                       80: //Check which conveyor
                           //Popup 2 conveyor to popup conveyor 3
                           IF #Source_Location_Carousel.Device_Type = 16 AND #Destination_Location_Carousel.Device_Type = 17 AND "Control_DB".PopUp_Cnv[2].Cnv_Occupied AND
                               NOT "Control_DB".PopUp_Cnv[3].Cnv_Occupied AND "Control_DB".PopUp_Cnv[2].Inputs."Lift Down" AND "Control_DB".PopUp_Cnv[3].Inputs."Lift Down"
                           THEN //All good
                               "Control_DB"."Carrousel_Order Table".SM_State := "Control_DB".PopUp_Cnv[3].SM_State;
                               #State_Carrousel := 100;// Chain Transfer
                           ELSIF #Source_Location_Carousel.Device_Type = 16 AND #Destination_Location_Carousel.Device_Type = 17 AND "Control_DB".PopUp_Cnv[2].Cnv_Occupied AND
                               NOT "Control_DB".PopUp_Cnv[3].Cnv_Occupied AND (NOT "Control_DB".PopUp_Cnv[2].Inputs."Lift Down" OR NOT "Control_DB".PopUp_Cnv[3].Inputs."Lift Down")
                           THEN //Lift
                               "Control_DB"."Carrousel_Order Table".SM_State := "Control_DB".PopUp_Cnv[3].SM_State;
                               #State_Carrousel := 90;// Lift pop up 2 OR 3 
                           END_IF;

                       90:  //Lift PopUps
                               "Control_DB"."Carrousel_Order Table".SM_State := "Control_DB".PopUp_Cnv[3].SM_State;
                               "Control_DB".PopUp_Cnv[2].Instruction.Lift_Down := NOT "Control_DB".PopUp_Cnv[2].Running AND NOT "Control_DB".PopUp_Cnv[2].Inputs."Lift Down";
                               "Control_DB".PopUp_Cnv[3].Instruction.Lift_Down := NOT "Control_DB".PopUp_Cnv[3].Running AND NOT "Control_DB".PopUp_Cnv[3].Inputs."Lift Down";
                               IF "Control_DB".PopUp_Cnv[2].Inputs."Lift Down" AND "Control_DB".PopUp_Cnv[3].Inputs."Lift Down" THEN
                                   #State_Carrousel := 100;
                               END_IF;

                           100: //Start the transfer
                           //Popup 2 to popup 3 conveyors
                                   "Control_DB".PopUp_Cnv[2].Instruction.Transfer_To_ID := "Settings_DB".PopUp_Cnv_Settings[3].ID;
                               "Control_DB"."Carrousel_Order Table".SM_State := "Control_DB".PopUp_Cnv[3].SM_State;//Current machine state
                               "Control_DB".PopUp_Cnv[3].Instruction.Start_Transfer := NOT "Control_DB".PopUp_Cnv[3].Running;
                               "Control_DB".PopUp_Cnv[2].Instruction.Start_Transfer := NOT "Control_DB".PopUp_Cnv[2].Running;
                               IF "Control_DB".PopUp_Cnv[3].Running AND "Control_DB".PopUp_Cnv[2].Running THEN
                                   "Control_DB"."Carrousel_Order Table".Movement_Ready := TRUE;
                                   //"Control_DB"."Carrousel_Order Table".Task_Data_Available := FALSE;
                                   #State_Carrousel := 110;
                               END_IF;

                       110: //Wait for the transfer to complete
                           //Popup 2 to popup 3 conveyors
                           "Control_DB"."Carrousel_Order Table".SM_State := "Control_DB".PopUp_Cnv[3].SM_State;
                           IF "Control_DB".PopUp_Cnv[3].Done AND "Control_DB".PopUp_Cnv[2].Done
                           THEN
                               "Control_DB"."Carrousel_Order Table".Movement_Request_Complete := TRUE;
                               #State_Carrousel := 120;
                           END_IF;

                       120: //Wait for the ACK before we go back to Idle
                           "Control_DB"."Carrousel_Order Table".SM_State := "Control_DB".PopUp_Cnv[3].SM_State;
                           IF "Control_DB"."Carrousel_Order Table".Movement_Request_Complete_Ack THEN
                               #State_Carrousel := 250;
                           END_IF;

                           //=========================== Transfer to pick station (From Pop Conveyor 4)  ===========================

                       130: //Check which conveyor
                               //Pop conveyor 4 to popup conveyor 1 (Pick Station)    
                           IF #Source_Location_Carousel.Device_Type = 18 AND #Destination_Location_Carousel.Device_Type = 41 AND "Control_DB".PopUp_Cnv[4].Cnv_Occupied AND
                               "Pick Station" AND "Control_DB".PopUp_Cnv[4].Inputs."Lift Down" AND "Control_DB".PopUp_Cnv[1].Inputs."Lift Down"
                           THEN //All good
                               "Control_DB"."Carrousel_Order Table".SM_State := "Control_DB".PopUp_Cnv[1].SM_State;
                               #State_Carrousel := 150;// Chain Transfer
                           ELSIF #Source_Location_Carousel.Device_Type = 18 AND #Destination_Location_Carousel.Device_Type = 41 AND "Control_DB".PopUp_Cnv[4].Cnv_Occupied AND
                               "Pick Station" AND (NOT "Control_DB".PopUp_Cnv[4].Inputs."Lift Down" OR NOT "Control_DB".PopUp_Cnv[1].Inputs."Lift Down")
                           THEN //Lift
                               "Control_DB"."Carrousel_Order Table".SM_State := "Control_DB".PopUp_Cnv[1].SM_State;
                               #State_Carrousel := 140;// Lift pop up 1
                           END_IF;

                       140:  //Lift PopUp
                           "Control_DB"."Carrousel_Order Table".SM_State := "Control_DB".PopUp_Cnv[1].SM_State;
                            // "Control_DB".PopUp_Cnv[1].Instruction.Lift_Down := NOT "Control_DB".PopUp_Cnv[1].Running AND NOT "Control_DB".PopUp_Cnv[1].Inputs."Lift Down";
                            "Control_DB".PopUp_Cnv[4].Instruction.Lift_Down := NOT "Control_DB".PopUp_Cnv[4].Running AND NOT "Control_DB".PopUp_Cnv[4].Inputs."Lift Down" ;
                            IF (*"Control_DB".PopUp_Cnv[1].Inputs."Lift Down" AND*) "Control_DB".PopUp_Cnv[4].Inputs."Lift Down" THEN
                                   #State_Carrousel := 150;
                               END_IF;

                       150: //Start the transfer
                           //Popup 4 TO Pick station conveyors
                               "Control_DB"."Carrousel_Order Table".SM_State := "Control_DB".PopUp_Cnv[1].SM_State;//Current machine state
                               "Control_DB".PopUp_Cnv[1].Instruction.Start_Transfer := NOT "Control_DB".PopUp_Cnv[1].Running;
                               IF "Control_DB".PopUp_Cnv[1].Running THEN
                                   "Control_DB"."Carrousel_Order Table".Movement_Ready := TRUE;
                                  // "Control_DB"."Carrousel_Order Table".Task_Data_Available := FALSE;
                                   #State_Carrousel := 160;
                               END_IF;

                       160: //Wait for the transfer to complete
                           //Popup 4 TO Pick station conveyors
                           "Control_DB"."Carrousel_Order Table".SM_State := "Control_DB".PopUp_Cnv[1].SM_State;
                           IF #Source_Location_Carousel.Device_Type = 18 AND #Destination_Location_Carousel.Device_Type = 41 AND
                               "Control_DB".PopUp_Cnv[1].Done
                           THEN
                               "Control_DB"."Carrousel_Order Table".Movement_Request_Complete := TRUE;
                               #State_Carrousel := 170;
                           END_IF;

                       170: //Wait for the ACK before we go back to Idle
                           "Control_DB"."Carrousel_Order Table".SM_State := "Control_DB".PopUp_Cnv[1].SM_State;
                           IF "Control_DB"."Carrousel_Order Table".Movement_Request_Complete_Ack THEN
                               #State_Carrousel := 250;
                           END_IF;

                           //=========================== Transfer from Pick station (To Pop Conveyor 1)  ===========================

                       180: //Check which conveyor
                               //Pick to popup conveyor 1   
                           IF #Source_Location_Carousel.Device_Type = 41 AND #Destination_Location_Carousel.Device_Type = 15 AND NOT "Pick Station" AND
                               NOT "Control_DB".PopUp_Cnv[1].Cnv_Occupied AND "Control_DB".PopUp_Cnv[1].Inputs."Lift Down"
                           THEN //All good
                               "Control_DB"."Carrousel_Order Table".SM_State := "Control_DB".PopUp_Cnv[1].SM_State;
                               #State_Carrousel := 200;// Chain Transfer
                           ELSIF #Source_Location_Carousel.Device_Type = 41 AND #Destination_Location_Carousel.Device_Type = 15 AND NOT "Pick Station" AND
                               NOT "Control_DB".PopUp_Cnv[1].Cnv_Occupied AND NOT "Control_DB".PopUp_Cnv[1].Inputs."Lift Down"
                           THEN //Lift
                               "Control_DB"."Carrousel_Order Table".SM_State := "Control_DB".PopUp_Cnv[1].SM_State;
                               #State_Carrousel := 190;// Lift pop up 1
                           END_IF;

                       190:  //Lift PopUps
                           "Control_DB"."Carrousel_Order Table".SM_State := "Control_DB".PopUp_Cnv[1].SM_State;
                           "Control_DB".PopUp_Cnv[1].Instruction.Lift_Down := NOT "Control_DB".PopUp_Cnv[1].Running AND NOT "Control_DB".PopUp_Cnv[1].Inputs."Lift Down";
                           IF "Control_DB".PopUp_Cnv[1].Inputs."Lift Down" THEN
                               #State_Carrousel := 200;
                           END_IF;

                       200: //Start the transfer
                           //Pick station TO Popup 1 conveyors
                               "Control_DB"."Carrousel_Order Table".SM_State := "Control_DB".PopUp_Cnv[1].SM_State;//Current machine state
                               "Control_DB".PopUp_Cnv[1].Instruction.Start_Transfer := NOT "Control_DB".PopUp_Cnv[1].Running;
                               IF "Control_DB".PopUp_Cnv[1].Running AND NOT "Control_DB".PopUp_Cnv[1].Done THEN
                                   "Control_DB"."Carrousel_Order Table".Movement_Ready := TRUE;
                                   //"Control_DB"."Carrousel_Order Table".Task_Data_Available := FALSE;
                                   #State_Carrousel := 210;
                               END_IF;

                       210: //Wait for the transfer to complete
                           //Pick station TO PopUp 1 conveyors
                           "Control_DB"."Carrousel_Order Table".SM_State := "Control_DB".PopUp_Cnv[1].SM_State;
                           IF "Control_DB".PopUp_Cnv[1].Done THEN
                               "Control_DB"."Carrousel_Order Table".Movement_Request_Complete := TRUE;
                               #State_Carrousel := 220;
                           END_IF;

                       220: //Wait for the ACK before we go back to Idle
                           "Control_DB"."Carrousel_Order Table".SM_State := "Control_DB".PopUp_Cnv[1].SM_State;
                           IF "Control_DB"."Carrousel_Order Table".Movement_Request_Complete_Ack THEN
                               #State_Carrousel := 250;
                           END_IF;

                           //=========================== Weigh Pallet  ===========================
                       230:
                          // "Control_DB"."Carrousel_Order Table".Task_Data_Available := FALSE;
                           "Control_DB"."Weighing Station".Start := TRUE;
                           "Control_DB"."Carrousel_Order Table".Movement_Ready := TRUE;
                           "Control_DB"."Carrousel_Order Table".SM_State := INT_TO_UINT("State_WS");
                           //Lift PopUp 1
                           "Control_DB".PopUp_Cnv[1].Instruction.Lift_Up := NOT "Control_DB".PopUp_Cnv[1].Running AND NOT "Control_DB".PopUp_Cnv[1].Inputs."Lift Up";

                           "IEC_Timer_0_DB_9".TON(IN:="Control_DB".PopUp_Cnv[1].Inputs."Lift Up",
                                                  PT:=T#500MS);
                           IF "IEC_Timer_0_DB_9".Q THEN
                               "Control_DB"."Weighing Station".Start := fALSE;
                               "IEC_Timer_0_DB_9".TON(IN := fALSE,
                                                      PT := T#0MS);
                               #State_Carrousel := 232;
                           END_IF;

                       232:
                           "Control_DB"."Carrousel_Order Table".SM_State := INT_TO_UINT("State_WS");
                           IF "Control_DB"."Weighing Station".Done THEN
                               "Control_DB"."Carrousel_Order Table".Movement_Request_Complete := TRUE;
                               IF "Control_DB"."Carrousel_Order Table".Movement_Request_Complete_Ack THEN
                                   #State_Carrousel := 250;
                               END_IF;
                           ELSE
                               #State_Carrousel := 250;
                           END_IF;

                           //=========================== Reset and Error States ===========================
                           250: //Reset all variable and return to idle

                           //Reset the OPC control variables
                               "Control_DB"."Carrousel_Order Table".SM_State := 0;
                               "Control_DB"."Carrousel_Order Table".Movement_Ready := FALSE;
                               "Control_DB"."Carrousel_Order Table".Movement_Request_Complete := FALSE;
                               "Control_DB"."Carrousel_Order Table".Movement_Request_Complete_Ack := FALSE;
                               "Control_DB"."Carrousel_Order Table".Task_Metadata := '';

                               "Control_DB"."Carrousel_Order Table".Task_Data_Available := FALSE; // Send the Task Data Available from WCS 
                               "Control_DB"."Carrousel_Order Table".Task_Type := 0; //  Send the Task Type - Roller to Roller Conveyor = Task Type = 6
                               "Control_DB"."Carrousel_Order Table".Task_ID := 0; // Send the Task ID number;
                               "Control_DB"."Carrousel_Order Table".Source_Location := 0; // Send the Source Location from the Conveyor
                               "Control_DB"."Carrousel_Order Table".Destination_Location := 0; // Send the Destination Location 
                               #Destination_Location_Carousel.Device_Type:=0;
                               #Source_Location_Carousel.Device_Type := 0;

                           //Reset conveyor variables
                           "Control_DB".Inbound_Cnv.Instruction.Start_Transfer := FALSE;
                           "Control_DB".Inbound_Cnv.Instruction.Task_ID := 0;
                           "Control_DB".Inbound_Cnv.Instruction.Task_Metadata := '';
                           "Control_DB".Inbound_Cnv.Current_Task_Type := 0;
                           "Control_DB".Inbound_Cnv.Instruction.Transfer_From_ID := 0;
                           "Control_DB".Inbound_Cnv.Instruction.Transfer_To_ID := 0;

                           "Control_DB".Outbound_Cnv.Instruction.Start_Transfer := FALSE;
                           "Control_DB".Outbound_Cnv.Instruction.Task_ID := 0;
                           "Control_DB".Outbound_Cnv.Instruction.Task_Metadata := '';
                           "Control_DB".Outbound_Cnv.Current_Task_Type := 0;
                           "Control_DB".Outbound_Cnv.Instruction.Transfer_From_ID := 0;
                           "Control_DB".Outbound_Cnv.Instruction.Transfer_To_ID := 0;

                           FOR #i := 1 TO 4 DO
                               "Control_DB".PopUp_Cnv[#i].Instruction.Start_Transfer := FALSE;
                               "Control_DB".PopUp_Cnv[#i].Instruction.Task_ID := 0;
                               "Control_DB".PopUp_Cnv[#i].Instruction.Task_Metadata := '';
                               "Control_DB".PopUp_Cnv[#i].Current_Task_Type := 0;
                               "Control_DB".PopUp_Cnv[#i].Instruction.Transfer_From_ID := 0;
                               "Control_DB".PopUp_Cnv[#i].Instruction.Transfer_To_ID := 0;
                           END_FOR;

                           "Error_Word_1".%X1 := FALSE;

                           #State_Carrousel := 0;

                           400:// Error state
                               "Control_DB"."Carrousel_Order Table".Task_Metadata := '';
                               "Control_DB"."Carrousel_Order Table".Task_Data_Available := FALSE; // Send the Task Data Available from WCS 
                               "Control_DB"."Carrousel_Order Table".Task_Type := 0; //  Send the Task Type - Roller to Roller Conveyor = Task Type = 6
                               "Control_DB"."Carrousel_Order Table".Task_ID := 0; // Send the Task ID number;
                               "Control_DB"."Carrousel_Order Table".Source_Location := 0; // Send the Source Location from the Conveyor
                               "Control_DB"."Carrousel_Order Table".Destination_Location := 0; // Send the Destination Location

                               #Destination_Location_Carousel.Device_Type := 0;
                               #Source_Location_Carousel.Device_Type := 0;


                           IF "Control_DB".VTD_Control.Instruction.Reset
                           THEN
                               #State_Carrousel := 250;
                           END_IF;

                       ELSE
                           ;
                   END_CASE;
                   ELSIF "Carrousel_In_Automatic" AND NOT #OPC_Enable THEN
                       "Control_DB"."Carrousel_Order Table".Task_Metadata := '';
                       //Reset all variable and return to idle

                       //Reset the OPC control variables
                       "Control_DB"."Carrousel_Order Table".SM_State := 0;
                       "Control_DB"."Carrousel_Order Table".Movement_Ready := FALSE;
                       "Control_DB"."Carrousel_Order Table".Movement_Request_Complete := FALSE;

                       "Control_DB"."Carrousel_Order Table".Task_Data_Available := FALSE; // Send the Task Data Available from WCS 
                       "Control_DB"."Carrousel_Order Table".Task_Type := 0; //  Send the Task Type - Roller to Roller Conveyor = Task Type = 6
                       "Control_DB"."Carrousel_Order Table".Task_ID := 0; // Send the Task ID number;
                       "Control_DB"."Carrousel_Order Table".Source_Location := 0; // Send the Source Location from the Conveyor
                       "Control_DB"."Carrousel_Order Table".Destination_Location := 0; // Send the Destination Location

                       #Destination_Location_Carousel.Device_Type := 0;
                       #Source_Location_Carousel.Device_Type := 0;

                       //Reset conveyor variables
                       "Control_DB".Inbound_Cnv.Instruction.Start_Transfer := FALSE;
                       "Control_DB".Inbound_Cnv.Instruction.Task_ID := 0;
                       "Control_DB".Inbound_Cnv.Instruction.Task_Metadata := '';//
                       "Control_DB".Inbound_Cnv.Instruction.Transfer_From_ID := 0;
                       "Control_DB".Inbound_Cnv.Instruction.Transfer_To_ID := 0;

                       "Control_DB".Outbound_Cnv.Instruction.Start_Transfer := FALSE;
                       "Control_DB".Outbound_Cnv.Instruction.Task_ID := 0;
                       "Control_DB".Outbound_Cnv.Instruction.Task_Metadata := '';//
                       "Control_DB".Outbound_Cnv.Instruction.Transfer_From_ID := 0;
                       "Control_DB".Outbound_Cnv.Instruction.Transfer_To_ID := 0;

                       FOR #i := 1 TO 4 DO
                           "Control_DB".PopUp_Cnv[#i].Instruction.Start_Transfer := FALSE;
                           "Control_DB".PopUp_Cnv[#i].Instruction.Task_ID := 0;
                           "Control_DB".PopUp_Cnv[#i].Instruction.Task_Metadata := '';
                           "Control_DB".PopUp_Cnv[#i].Current_Task_Type := 0;
                           "Control_DB".PopUp_Cnv[#i].Instruction.Transfer_From_ID := 0;
                           "Control_DB".PopUp_Cnv[#i].Instruction.Transfer_To_ID := 0;
                       END_FOR;
                   END_IF;
       END_REGION
   END_REGION

   REGION SHUTTLES POSITION
       FOR #f := 1 TO "Settings_DB".System_Settings.Shuttle_Count DO
           "Control_DB".Shuttles_Position[#f].x := "Shuttle_MQTT_DB".Shuttle_MQTT[#f].Message.Shuttle_Status.Position_X;
           "Control_DB".Shuttles_Position[#f].y := "Shuttle_MQTT_DB".Shuttle_MQTT[#f].Message.Shuttle_Status.Position_Y;
       END_FOR;
   END_REGION

   REGION SM STATE MAESTRO
       // Statement section - Send the State machine to Maestro "Emulating" openTCS states
       // 
      // // "Control_DB".WMS_OPC_UA.SM_State_Maestro; // State to send Devices to Maestro
      //  IF #State_VTD = 0 THEN

      //      "Control_DB"."VTD_Order Table".SM_State_Maestro := 0;//"LIMBO" condition 

      //  ELSIF "Control_DB"."VTD_Order Table".SM_State = 10 THEN
      //      ;
      //      // "Control_DB".WMS_OPC_UA.SM_State_Maestro := 1;//RAW conidtion => Maestro will write this condition

      //      //////////////////////////////////////////////////////////////////////////////////////////////////////////////////////      
      //      // QUEUED ANY DEVICE    
      //  // ELSIF "Control_DB".WMS_OPC_UA.Task_Data_Available AND #State >= 10 AND #State <= 20 THEN
      //  ELSIF "Control_DB"."VTD_Order Table".Task_Data_Available AND NOT "Control_DB"."VTD_Order Table".Movement_Ready AND "Control_DB"."VTD_Order Table".SM_State_Maestro = 1 THEN
      //      "Control_DB"."VTD_Order Table".SM_State_Maestro := 2;//QUEUED condition =>ANY device (Conveyor, VTD OR Shuttle)  

      //      //////////////////////////////////////////////////////////////////////////////////////////////////////////////////////       
      //      // Any Device RUNNING on the system (VTD - Conveyor Transfer - Shuttle Transfer) 
      //  ELSIF ("Control_DB"."VTD_Order Table".Task_Type = 4 OR "Control_DB"."VTD_Order Table".Task_Type = 5
      //      OR "Control_DB"."VTD_Order Table".Task_Type = 1 OR "Control_DB"."VTD_Order Table".Task_Type = 2 OR "Control_DB"."VTD_Order Table".Task_Type = 3)
      //      AND "Control_DB"."VTD_Order Table".Movement_Ready AND NOT "Control_DB"."VTD_Order Table".Movement_Request_Complete THEN

      //      "Control_DB"."VTD_Order Table".SM_State_Maestro := 3;//RUNNING condition

      //      // Any Device DONE on the system (VTD - Coneveyor Transfer - Shuttle Transfer) 
      //  ELSIF ("Control_DB"."VTD_Order Table".Task_Type = 4 OR "Control_DB"."VTD_Order Table".Task_Type = 5
      //      OR "Control_DB"."VTD_Order Table".Task_Type = 1 OR "Control_DB"."VTD_Order Table".Task_Type = 2 OR "Control_DB"."VTD_Order Table".Task_Type = 3)
      //      AND (*"Control_DB".WMS_OPC_UA.Movement_Request_Complete AND "Control_DB".WMS_OPC_UA.Movement_Ready*)#State_VTD = 120 OR #State_VTD = 45 OR #State_VTD = 90 THEN

      //      "Control_DB"."VTD_Order Table".SM_State_Maestro := 4;//DONE condition

      //      // Any Device ERRORS on the system (VTD - Coneveyor Transfer - Shuttle Transfer)  
      //  ELSIF ("Control_DB"."VTD_Order Table".Task_Type = 4 OR "Control_DB"."VTD_Order Table".Task_Type = 5
      //      OR "Control_DB"."VTD_Order Table".Task_Type = 1 OR "Control_DB"."VTD_Order Table".Task_Type = 2 OR "Control_DB"."VTD_Order Table".Task_Type = 3)
      //      AND "Control_DB"."VTD_Order Table".SM_State = 400 THEN

      //      "Control_DB"."VTD_Order Table".SM_State_Maestro := 5;//ERROR condition => Conveyors   
      //  END_IF;
      //      /////////////////////////////////////////////////////////////////////////////////////////////        



       // "Control_DB".WMS_OPC_UA.SM_State_Maestro; // State to send Devices to Maestro
        IF #State_VTD = 0 THEN
            ;
            //"System_DB_VTD".OrderTable[1].OPC_Control.SM_State_Maestro := 0;//"LIMBO" condition 

        ELSIF "Control_DB"."VTD_Order Table".SM_State = 10 THEN
            ;
            // "Control_DB".WMS_OPC_UA.SM_State_Maestro := 1;//RAW conidtion => Maestro will write this condition

            //////////////////////////////////////////////////////////////////////////////////////////////////////////////////////      
            // QUEUED ANY DEVICE    
        // ELSIF "Control_DB".WMS_OPC_UA.Task_Data_Available AND #State >= 10 AND #State <= 20 THEN
        ELSIF "Control_DB"."VTD_Order Table".Task_Data_Available AND NOT "Control_DB"."VTD_Order Table".Movement_Ready AND "System_DB_VTD".OrderTable[1].OPC_Control.SM_State_Maestro = 1 THEN
            "System_DB_VTD".OrderTable[1].OPC_Control.SM_State_Maestro := 2;//QUEUED condition =>ANY device (Conveyor, VTD OR Shuttle)  

            //////////////////////////////////////////////////////////////////////////////////////////////////////////////////////       
            // Any Device RUNNING on the system (VTD - Conveyor Transfer - Shuttle Transfer) 
        ELSIF ("Control_DB"."VTD_Order Table".Task_Type = 4 OR "Control_DB"."VTD_Order Table".Task_Type = 5
            OR "Control_DB"."VTD_Order Table".Task_Type = 1 OR "Control_DB"."VTD_Order Table".Task_Type = 2 OR "Control_DB"."VTD_Order Table".Task_Type = 3)
            AND "Control_DB"."VTD_Order Table".Movement_Ready AND NOT "Control_DB"."VTD_Order Table".Movement_Request_Complete THEN

            "System_DB_VTD".OrderTable[1].OPC_Control.SM_State_Maestro  := 3;//RUNNING condition

            // Any Device DONE on the system (VTD - Coneveyor Transfer - Shuttle Transfer) 
        ELSIF ("Control_DB"."VTD_Order Table".Task_Type = 4 OR "Control_DB"."VTD_Order Table".Task_Type = 5
            OR "Control_DB"."VTD_Order Table".Task_Type = 1 OR "Control_DB"."VTD_Order Table".Task_Type = 2 OR "Control_DB"."VTD_Order Table".Task_Type = 3)
            AND (*"Control_DB".WMS_OPC_UA.Movement_Request_Complete AND "Control_DB".WMS_OPC_UA.Movement_Ready*)#State_VTD = 120 OR #State_VTD = 45 OR #State_VTD = 90 THEN

            "System_DB_VTD".OrderTable[1].OPC_Control.SM_State_Maestro := 4;//DONE condition

            // Any Device ERRORS on the system (VTD - Coneveyor Transfer - Shuttle Transfer)  
        ELSIF ("Control_DB"."VTD_Order Table".Task_Type = 4 OR "Control_DB"."VTD_Order Table".Task_Type = 5
            OR "Control_DB"."VTD_Order Table".Task_Type = 1 OR "Control_DB"."VTD_Order Table".Task_Type = 2 OR "Control_DB"."VTD_Order Table".Task_Type = 3)
            AND "Control_DB"."VTD_Order Table".SM_State = 400 THEN

            "System_DB_VTD".OrderTable[1].OPC_Control.SM_State_Maestro := 5;//ERROR condition => Conveyors   
        END_IF;
            /////////////////////////////////////////////////////////////////////////////////////////////        


      //  //     //////////////////////////////////////////////////////////////////////////////////////////////////////////////////////       
      //  //     // Any VTD RUNNING on the system (VTD) 
      //  // ELSIF "Control_DB".WMS_OPC_UA.Task_Type = 1
      //  //     AND "Control_DB".WMS_OPC_UA.SM_State >= 35 AND "Control_DB".WMS_OPC_UA.SM_State < 100 AND #State > 20 THEN

      //  //     "Control_DB".WMS_OPC_UA.SM_State_Maestro := 3;//RUNNING condition => VTD

      //  //     // Any VTD DONE on the system (VTD) 
      //  // ELSIF "Control_DB".WMS_OPC_UA.Task_Type = 1
      //  //     AND "Control_DB".WMS_OPC_UA.SM_State = 100 AND #State > 20 THEN

      //  //     "Control_DB".WMS_OPC_UA.SM_State_Maestro := 4;//DONE condition => VTD

      //  //     // Any VTD ERRORS on the system (VTD) 
      //  // ELSIF "Control_DB".WMS_OPC_UA.Task_Type = 1
      //  //     AND "Control_DB".WMS_OPC_UA.SM_State = 400 THEN

      //  //     "Control_DB".WMS_OPC_UA.SM_State_Maestro := 5;//ERROR condition => VTD   



      //  //     //////////////////////////////////////////////////////////////////////////////////////////////////////////////////////       
      //  //     // Any Shuttle Interlock RUNNING on the system (Shuttle) 
      //  // ELSIF "Control_DB".WMS_OPC_UA.Task_Type = 2 OR "Control_DB".WMS_OPC_UA.Task_Type = 3
      //  //     AND "Control_DB".WMS_OPC_UA.SM_State >= 35 AND "Control_DB".WMS_OPC_UA.SM_State < 100 AND #State > 20 THEN

      //  //     "Control_DB".WMS_OPC_UA.SM_State_Maestro := 3;//RUNNING condition => Shuttle

      //  //     // Any Shuttle Interlock  DONE on the system (Shuttle) 
      //  // ELSIF "Control_DB".WMS_OPC_UA.Task_Type = 2 OR "Control_DB".WMS_OPC_UA.Task_Type = 3
      //  //     AND "Control_DB".WMS_OPC_UA.SM_State = 100 AND #State > 20 THEN

      //  //     "Control_DB".WMS_OPC_UA.SM_State_Maestro := 4;//DONE condition => Shuttle

      //  //     // Any Shuttle Interlock ERRORS on the system (Shuttle) 
      //  // ELSIF "Control_DB".WMS_OPC_UA.Task_Type = 2 OR "Control_DB".WMS_OPC_UA.Task_Type = 3
      //  //     AND "Control_DB".WMS_OPC_UA.SM_State = 400 THEN

      //  //     "Control_DB".WMS_OPC_UA.SM_State_Maestro := 5;//ERROR condition => Shuttle          

      //  // END_IF;


       // // "Control_DB".WMS_OPC_UA.SM_State_Maestro; // State to send Devices to Maestro
       //  IF #State_VTD = 0 THEN

       //      "Control_DB"."VTD_Order Table".SM_State_Maestro := 0;//"LIMBO" condition 

       //  ELSIF "Control_DB"."VTD_Order Table".SM_State = 10 THEN
       //      ;
       //      // "Control_DB".WMS_OPC_UA.SM_State_Maestro := 1;//RAW conidtion => Maestro will write this condition

       //      //////////////////////////////////////////////////////////////////////////////////////////////////////////////////////      
       //      // QUEUED ANY DEVICE    
       //  // ELSIF "Control_DB".WMS_OPC_UA.Task_Data_Available AND #State >= 10 AND #State <= 20 THEN
       //  ELSIF "Control_DB"."VTD_Order Table".Task_Data_Available AND NOT "Control_DB"."VTD_Order Table".Movement_Ready AND "Control_DB"."VTD_Order Table".SM_State_Maestro = 1 THEN
       //      "Control_DB"."VTD_Order Table".SM_State_Maestro := 2;//QUEUED condition =>ANY device (Conveyor, VTD OR Shuttle)  

       //      //////////////////////////////////////////////////////////////////////////////////////////////////////////////////////       
       //      // Any Device RUNNING on the system (VTD - Conveyor Transfer - Shuttle Transfer) 
       //  ELSIF ("Control_DB"."VTD_Order Table".Task_Type = 4 OR "Control_DB"."VTD_Order Table".Task_Type = 5
       //      OR "Control_DB"."VTD_Order Table".Task_Type = 1 OR "Control_DB"."VTD_Order Table".Task_Type = 2 OR "Control_DB"."VTD_Order Table".Task_Type = 3)
       //      AND "Control_DB"."VTD_Order Table".Movement_Ready AND NOT "Control_DB"."VTD_Order Table".Movement_Request_Complete THEN

       //      "Control_DB"."VTD_Order Table".SM_State_Maestro := 3;//RUNNING condition

       //      // Any Device DONE on the system (VTD - Coneveyor Transfer - Shuttle Transfer) 
       //  ELSIF ("Control_DB"."VTD_Order Table".Task_Type = 4 OR "Control_DB"."VTD_Order Table".Task_Type = 5
       //      OR "Control_DB"."VTD_Order Table".Task_Type = 1 OR "Control_DB"."VTD_Order Table".Task_Type = 2 OR "Control_DB"."VTD_Order Table".Task_Type = 3)
       //      AND (*"Control_DB".WMS_OPC_UA.Movement_Request_Complete AND "Control_DB".WMS_OPC_UA.Movement_Ready*)#State_VTD = 120 OR #State_VTD = 45 OR #State_VTD = 90 THEN

       //      "Control_DB"."VTD_Order Table".SM_State_Maestro := 4;//DONE condition

       //      // Any Device ERRORS on the system (VTD - Coneveyor Transfer - Shuttle Transfer)  
       //  ELSIF ("Control_DB"."VTD_Order Table".Task_Type = 4 OR "Control_DB"."VTD_Order Table".Task_Type = 5
       //      OR "Control_DB"."VTD_Order Table".Task_Type = 1 OR "Control_DB"."VTD_Order Table".Task_Type = 2 OR "Control_DB"."VTD_Order Table".Task_Type = 3)
       //      AND "Control_DB"."VTD_Order Table".SM_State = 400 THEN

       //      "Control_DB"."VTD_Order Table".SM_State_Maestro := 5;//ERROR condition => Conveyors   
       //  END_IF;
       //      /////////////////////////////////////////////////////////////////////////////////////////////        

       //  //     //////////////////////////////////////////////////////////////////////////////////////////////////////////////////////       
       //  //     // Any VTD RUNNING on the system (VTD) 
       //  // ELSIF "Control_DB".WMS_OPC_UA.Task_Type = 1
       //  //     AND "Control_DB".WMS_OPC_UA.SM_State >= 35 AND "Control_DB".WMS_OPC_UA.SM_State < 100 AND #State > 20 THEN

       //  //     "Control_DB".WMS_OPC_UA.SM_State_Maestro := 3;//RUNNING condition => VTD

       //  //     // Any VTD DONE on the system (VTD) 
       //  // ELSIF "Control_DB".WMS_OPC_UA.Task_Type = 1
       //  //     AND "Control_DB".WMS_OPC_UA.SM_State = 100 AND #State > 20 THEN

       //  //     "Control_DB".WMS_OPC_UA.SM_State_Maestro := 4;//DONE condition => VTD

       //  //     // Any VTD ERRORS on the system (VTD) 
       //  // ELSIF "Control_DB".WMS_OPC_UA.Task_Type = 1
       //  //     AND "Control_DB".WMS_OPC_UA.SM_State = 400 THEN

       //  //     "Control_DB".WMS_OPC_UA.SM_State_Maestro := 5;//ERROR condition => VTD   



       //  //     //////////////////////////////////////////////////////////////////////////////////////////////////////////////////////       
       //  //     // Any Shuttle Interlock RUNNING on the system (Shuttle) 
       //  // ELSIF "Control_DB".WMS_OPC_UA.Task_Type = 2 OR "Control_DB".WMS_OPC_UA.Task_Type = 3
       //  //     AND "Control_DB".WMS_OPC_UA.SM_State >= 35 AND "Control_DB".WMS_OPC_UA.SM_State < 100 AND #State > 20 THEN

       //  //     "Control_DB".WMS_OPC_UA.SM_State_Maestro := 3;//RUNNING condition => Shuttle

       //  //     // Any Shuttle Interlock  DONE on the system (Shuttle) 
       //  // ELSIF "Control_DB".WMS_OPC_UA.Task_Type = 2 OR "Control_DB".WMS_OPC_UA.Task_Type = 3
       //  //     AND "Control_DB".WMS_OPC_UA.SM_State = 100 AND #State > 20 THEN

       //  //     "Control_DB".WMS_OPC_UA.SM_State_Maestro := 4;//DONE condition => Shuttle

       //  //     // Any Shuttle Interlock ERRORS on the system (Shuttle) 
       //  // ELSIF "Control_DB".WMS_OPC_UA.Task_Type = 2 OR "Control_DB".WMS_OPC_UA.Task_Type = 3
       //  //     AND "Control_DB".WMS_OPC_UA.SM_State = 400 THEN

       //  //     "Control_DB".WMS_OPC_UA.SM_State_Maestro := 5;//ERROR condition => Shuttle          

       //  // END_IF;

   END_REGION


   REGION SM STATE MAESTRO - Carousel
       // Statement section - Send the State machine to Maestro "Emulating" openTCS states
       // 

       (*
       IF #State_Carrousel = 0 THEN

           "Control_DB"."Carrousel_Order Table".SM_State_Maestro := 0;//"LIMBO" condition 

       ELSIF "Control_DB"."Carrousel_Order Table".SM_State = 10 THEN
           ;
           // "Control_DB".WMS_OPC_UA.SM_State_Maestro := 1;//RAW conidtion => Maestro will write this condition

           //////////////////////////////////////////////////////////////////////////////////////////////////////////////////////      
           // QUEUED ANY DEVICE    
           // ELSIF "Control_DB".WMS_OPC_UA.Task_Data_Available AND #State >= 10 AND #State <= 20 THEN
       ELSIF "Control_DB"."Carrousel_Order Table".Task_Data_Available AND NOT "Control_DB"."Carrousel_Order Table".Movement_Ready AND "Control_DB"."Carrousel_Order Table".SM_State_Maestro = 1 THEN
           "Control_DB"."Carrousel_Order Table".SM_State_Maestro := 2;//QUEUED condition =>ANY device (Conveyor, VTD OR Shuttle)  

           //////////////////////////////////////////////////////////////////////////////////////////////////////////////////////       
           // Any Device RUNNING on the system (VTD - Conveyor Transfer - Shuttle Transfer) 
       ELSIF ("Control_DB"."Carrousel_Order Table".Task_Type = 6 OR "Control_DB"."Carrousel_Order Table".Task_Type = 7
           OR "Control_DB"."Carrousel_Order Table".Task_Type = 8 OR "Control_DB"."Carrousel_Order Table".Task_Type = 9
           OR "Control_DB"."Carrousel_Order Table".Task_Type = 10 OR "Control_DB"."Carrousel_Order Table".Task_Type = 14 OR "Control_DB"."Carrousel_Order Table".Task_Type = 16)
           AND "Control_DB"."Carrousel_Order Table".Movement_Ready AND NOT "Control_DB"."Carrousel_Order Table".Movement_Request_Complete THEN

           "Control_DB"."Carrousel_Order Table".SM_State_Maestro := 3;//RUNNING condition

           // Any Device DONE on the system (VTD - Coneveyor Transfer - Shuttle Transfer) 
       ELSIF ("Control_DB"."Carrousel_Order Table".Task_Type = 6 OR "Control_DB"."Carrousel_Order Table".Task_Type = 7
           OR "Control_DB"."Carrousel_Order Table".Task_Type = 8 OR "Control_DB"."Carrousel_Order Table".Task_Type = 9
           OR "Control_DB"."Carrousel_Order Table".Task_Type = 10 OR "Control_DB"."Carrousel_Order Table".Task_Type = 14 OR "Control_DB"."Carrousel_Order Table".Task_Type = 16)
           AND (*"Control_DB".WMS_OPC_UA.Movement_Request_Complete AND "Control_DB".WMS_OPC_UA.Movement_Ready*)#State_Carrousel = 70 OR #State_Carrousel = 120 OR #State_Carrousel = 170 OR #State_Carrousel = 220 OR #State_Carrousel = 232 THEN

           "Control_DB"."Carrousel_Order Table".SM_State_Maestro := 4;//DONE condition

           // Any Device ERRORS on the system (VTD - Coneveyor Transfer - Shuttle Transfer)  
       ELSIF ("Control_DB"."Carrousel_Order Table".Task_Type = 6 OR "Control_DB"."Carrousel_Order Table".Task_Type = 7
           OR "Control_DB"."Carrousel_Order Table".Task_Type = 8 OR "Control_DB"."Carrousel_Order Table".Task_Type = 9
           OR "Control_DB"."Carrousel_Order Table".Task_Type = 10 OR "Control_DB"."Carrousel_Order Table".Task_Type = 14 OR "Control_DB"."Carrousel_Order Table".Task_Type = 16)
           AND "Control_DB"."Carrousel_Order Table".SM_State = 400 THEN

           "Control_DB"."Carrousel_Order Table".SM_State_Maestro := 5;//ERROR condition => Conveyors   
       END_IF;
       /////////////////////////////////////////////////////////////////////////////////////////////        
       *)


       IF #State_Carrousel = 0 THEN
           ;
           //"Control_DB"."Carrousel_Order Table".SM_State_Maestro := 0;//"LIMBO" condition 
           //"System_DB_Carousel".OrderTable[1].OPC_Control.SM_State_Maestro := 0;

       ELSIF "Control_DB"."Carrousel_Order Table".SM_State = 10 THEN
           ;
           // "Control_DB".WMS_OPC_UA.SM_State_Maestro := 1;//RAW conidtion => Maestro will write this condition

           //////////////////////////////////////////////////////////////////////////////////////////////////////////////////////      
           // QUEUED ANY DEVICE    
           // ELSIF "Control_DB".WMS_OPC_UA.Task_Data_Available AND #State >= 10 AND #State <= 20 THEN
       ELSIF "Control_DB"."Carrousel_Order Table".Task_Data_Available AND NOT "Control_DB"."Carrousel_Order Table".Movement_Ready AND "System_DB_Carousel".OrderTable[1].OPC_Control.SM_State_Maestro = 1 THEN
           "System_DB_Carousel".OrderTable[1].OPC_Control.SM_State_Maestro := 2;//QUEUED condition =>ANY device (Conveyor, VTD OR Shuttle)  

           //////////////////////////////////////////////////////////////////////////////////////////////////////////////////////       
           // Any Device RUNNING on the system (VTD - Conveyor Transfer - Shuttle Transfer) 
       ELSIF ("Control_DB"."Carrousel_Order Table".Task_Type = 6 OR "Control_DB"."Carrousel_Order Table".Task_Type = 7
           OR "Control_DB"."Carrousel_Order Table".Task_Type = 8 OR "Control_DB"."Carrousel_Order Table".Task_Type = 9
           OR "Control_DB"."Carrousel_Order Table".Task_Type = 10 OR "Control_DB"."Carrousel_Order Table".Task_Type = 14 OR "Control_DB"."Carrousel_Order Table".Task_Type = 16)
           AND "Control_DB"."Carrousel_Order Table".Movement_Ready AND NOT "Control_DB"."Carrousel_Order Table".Movement_Request_Complete THEN

           "System_DB_Carousel".OrderTable[1].OPC_Control.SM_State_Maestro := 3;//RUNNING condition

           // Any Device DONE on the system (VTD - Coneveyor Transfer - Shuttle Transfer) 
       ELSIF ("Control_DB"."Carrousel_Order Table".Task_Type = 6 OR "Control_DB"."Carrousel_Order Table".Task_Type = 7
           OR "Control_DB"."Carrousel_Order Table".Task_Type = 8 OR "Control_DB"."Carrousel_Order Table".Task_Type = 9
           OR "Control_DB"."Carrousel_Order Table".Task_Type = 10 OR "Control_DB"."Carrousel_Order Table".Task_Type = 14 OR "Control_DB"."Carrousel_Order Table".Task_Type = 16)
           AND (*"Control_DB".WMS_OPC_UA.Movement_Request_Complete AND "Control_DB".WMS_OPC_UA.Movement_Ready*)#State_Carrousel = 70 OR #State_Carrousel = 120 OR #State_Carrousel = 170 OR #State_Carrousel = 220 OR #State_Carrousel = 232 THEN

           "System_DB_Carousel".OrderTable[1].OPC_Control.SM_State_Maestro := 4;//DONE condition

           // Any Device ERRORS on the system (VTD - Coneveyor Transfer - Shuttle Transfer)  
       ELSIF ("Control_DB"."Carrousel_Order Table".Task_Type = 6 OR "Control_DB"."Carrousel_Order Table".Task_Type = 7
           OR "Control_DB"."Carrousel_Order Table".Task_Type = 8 OR "Control_DB"."Carrousel_Order Table".Task_Type = 9
           OR "Control_DB"."Carrousel_Order Table".Task_Type = 10 OR "Control_DB"."Carrousel_Order Table".Task_Type = 14 OR "Control_DB"."Carrousel_Order Table".Task_Type = 16)
           AND "Control_DB"."Carrousel_Order Table".SM_State = 400 THEN

           "System_DB_Carousel".OrderTable[1].OPC_Control.SM_State_Maestro:= 5;//ERROR condition => Conveyors   
       END_IF;
       /////////////////////////////////////////////////////////////////////////////////////////////        





   END_REGION
END_FUNCTION_BLOCK

FUNCTION_BLOCK "Order_Table_FB_Carousel_1"   // FB34, SCL
{ S7_Optimized_Access := 'TRUE' }
VERSION : 0.1
// stored: AutoNumber true, IsIECCheckEnabled false, IsRetainMemResEnabled false, MemoryReserve 100, SetENOAutomatically false, UDAEnableTagReadback false
   VAR_INPUT
      System_Selected { ExternalWritable := 'False'} : Bool;
      AutoMan_Switch : Bool;   // Auto/Man Switch on CPU Panel - 1 = Auto, 0 = Manual
      CurrentTime { ExternalWritable := 'False'} : String;
      CurrentDTL : DTL;
      Watchdog : "Watchdog_Settings_UDT";
   END_VAR
   VAR_IN_OUT
      Cnv_Entry : "Inbound_Cnv_Control_UDT";
      Cnv_PopUp_1 : "PopUp_Cnv_Control";
      WeighingStation : "Stations_DB_UDT";
      ProfileStation : "Stations_DB_UDT";
      Cnv_PopUp_2 : "PopUp_Cnv_Control";
      Cnv_PopUp_3 : "PopUp_Cnv_Control";
      Cnv_PopUp_4 : "PopUp_Cnv_Control";
      Cnv_Exit : "Outbound_Cnv_Control";
      System : "System_UDT";
      Control_OPC_Ua : "WMS_OPC_UA";
   END_VAR
   VAR
      RTR_ITP1_CurrentOrder : UDInt;
      RTR_P1P2_CurrentOrder : UDInt;
      RTR_P3P4_CurrentOrder : UDInt;
      RTR_P4TO_CurrentOrder : UDInt;
      Roller_To_Roller_CurrentOrder : UDInt;
      Chain_To_Chain_CurrentOrder : UDInt;
      Pop4_To_PickSt_CurrentOrder : UDInt;
      PickSt_To_Pop1_CurrentOrder : UDInt;
      WeighingStation_CurrentOrder { ExternalWritable := 'False'} : UDInt := 0;
      ProfileStation_CurrentOrder { ExternalWritable := 'False'} : UDInt := 0;
      Roller_To_RollerDoneRTrig : R_TRIG;
      RTR_ITP1DoneRTrig { S7_SetPoint := 'True'} : R_TRIG;
      RTR_P1P2DoneRTrig { S7_SetPoint := 'True'} : R_TRIG;
      RTR_P3P4DoneRTrig { S7_SetPoint := 'True'} : R_TRIG;
      RTR_P4TODoneRTrig { S7_SetPoint := 'True'} : R_TRIG;
      Chain_To_ChainDoneRTrig : R_TRIG;
      Pop4_To_PickSt_DoneRTrig { S7_SetPoint := 'True'} : R_TRIG;
      PickSt_To_Pop1_DoneRTrig { S7_SetPoint := 'True'} : R_TRIG;
      WeighingStationDoneRTrig { ExternalWritable := 'False'} : R_TRIG;
      ProfileStationDoneRTrig { ExternalWritable := 'False'} : R_TRIG;
      PalletRefused_1_RTig { ExternalWritable := 'False'} : R_TRIG;
      ErrorRTrig { ExternalWritable := 'False'} : R_TRIG;
      CancelRTrig { ExternalWritable := 'False'} : R_TRIG;
      PauseRTrig { ExternalWritable := 'False'} : R_TRIG;
      ResumeRTrig { ExternalWritable := 'False'} : R_TRIG;
      Clear_Store : R_TRIG;
      Clear_Retrieve : R_TRIG;
      Canceling : Bool;
      RTR_ITP1_WatchdogTimer : TON_TIME;
      RTR_P1P2_WatchdogTimer : TON_TIME;
      RTR_P3P4_WatchdogTimer : TON_TIME;
      RTR_P4TO_WatchdogTimer : TON_TIME;
      Roller_To_Roller_WatchdogTimer { S7_SetPoint := 'True'} : TON_TIME;
      Chain_To_Chain_WatchdogTimer { S7_SetPoint := 'True'} : TON_TIME;
      Pop4_To_PickWatchdogTimer { S7_SetPoint := 'True'} : TON_TIME;
      PickSt_To_Pop1WatchdogTimer : TON_TIME;
      WeighingStation_WatchdogTimer : TON_TIME;
      ProfileStation_WatchdogTimer : TON_TIME;
      Roller_To_Roller_WatchdogStart { S7_SetPoint := 'True'} : Bool;
      RTR_ITP1_WatchdogStart : Bool;
      RTR_P1P2_WatchdogStart : Bool;
      RTR_P3P4_WatchdogStart : Bool;
      RTR_P4TO_WatchdogStart : Bool;
      Chain_To_Chain_WatchdogStart : Bool;
      Pop4_To_PickWatchdogStart : Bool;
      PickSt_To_Pop1WatchdogStart : Bool;
      WeighingStation_WatchdogStart : Bool;
      ProfileStation_WatchdogStart : Bool;
      dummy : Int;
      dummy_1 : Bool;
      dummy_3 : Bool;
   END_VAR
   VAR_TEMP
      i : DInt;
      n : DInt;
      EmptyOrder : "OrderTable_UDT";
      MaxRunningOrderNo : UInt;
   END_VAR
   VAR CONSTANT
      ROLLER_TO_ROLLER_DEVICE : String := 'Roller to Roller';
      CHAIN_TO_CHAIN_DEVICE : String := 'Chain to Chain';
      POP4_TO_PICK_DEVICE : String := 'Pop4 to Pick';
      PICK_TO_POP1_DEVICE : String := 'Pick to Pop1';
      WEIGH_STATION_DEVICE : String := 'Weigh Station';
      PROFILE_STATION_DEVICE : String := 'Profile Station';
      RUNNING_STATUS : String := 'Running';
      COMPLETED_STATUS : String := 'Completed';
      QUEUED_STATUS : String := 'Queued';
      PALLET_REFUSED_STATUS : String := 'Pallet Refused';
      ERROR_STATUS : String := 'Error';
      CANCELED_STATUS : String := 'Canceled';
      PAUSED_STATUS : String := 'Paused';
      ORDER_REFUSED : String := 'Refused';
      ERROR_CANCELED_STATUS : String := 'Error\Cancel';
   END_VAR
BEGIN

   // Converts the task type for strings 
   IF #System.OrderTable[1].OPC_Control.Task_Type = 6
       OR #System.OrderTable[1].OPC_Control.Task_Type =16
           OR #System.OrderTable[1].OPC_Control.Task_Type = 14 THEN // Roller to Roller OR Roller to Roller + Barcode scanner OR Roller To Roller + Profile Station 
       #System.OrderTable[1].Device := 'Roller to Roller';
   ELSIF #System.OrderTable[1].OPC_Control.Task_Type = 7 THEN
       #System.OrderTable[1].Device := 'Chain to Chain';
   ELSIF #System.OrderTable[1].OPC_Control.Task_Type = 8 THEN
       #System.OrderTable[1].Device := 'Pop4 to Pick';
   ELSIF #System.OrderTable[1].OPC_Control.Task_Type = 9 THEN
       #System.OrderTable[1].Device := 'Pick to Pop1' ;
   ELSIF #System.OrderTable[1].OPC_Control.Task_Type = 10 THEN
       #System.OrderTable[1].Device := 'Weigh Station';
   // ELSIF #System.OrderTable[1].OPC_Control.Task_Type = 14 THEN
   //     #System.OrderTable[1].Device := 'Profile Station';
   ELSE
       #System.OrderTable[1].Device := '';
   END_IF;


   REGION #New Order was Sent
       IF #System.OrderSent THEN
           //Count orders in Step Table
           FOR #i := 0 TO 20 DO
               IF #System.StepTable[#i].OrderNo <> 0
                   AND #System.StepTable[#i].StepNo <> 0
                   AND #System.StepTable[#i].PlaceTime <> ''
                   //AND #System.StepTable[#i].Device <> ''
                   AND #System.StepTable[#i].Status = #QUEUED_STATUS
               THEN
                   #n += 1;
               ELSE
                   EXIT;
               END_IF;
           END_FOR;

           IF #n > 0 THEN
               //shift order table down by Order number rows
               FOR #i := 99 TO (#n + 1) BY -1 DO
                   #System.OrderTable[#i] := #System.OrderTable[#i - #n];
               END_FOR;
               //copy data from step table to order table
               FOR #i := 0 TO #n DO
                   #System.OrderTable[#n - #i (*+ 1*)] := #System.StepTable[#i];
               END_FOR;
               //clean step table
               FOR #i := 0(*1*) TO 20 DO
                   #System.StepTable[#i] := #EmptyOrder;
               END_FOR;
               #System.CurrentOrder += #n;


               // Transfer Pallet Roller to Roller - 

               IF #Roller_To_Roller_CurrentOrder <> 0 THEN
                   #Roller_To_Roller_CurrentOrder += #n;
               END_IF;


               // Transfer Pallet Roller to Roller - Inbound to PP1

               IF #RTR_ITP1_CurrentOrder <> 0 THEN
                   #RTR_ITP1_CurrentOrder += #n;
               END_IF;

               // Transfer Pallet Roller to Roller - PP1 to PP2

               IF #RTR_P1P2_CurrentOrder <> 0 THEN
                   #RTR_P1P2_CurrentOrder += #n;
               END_IF;

               // Transfer Pallet Roller TO Roller - PP3 TO PP4

               IF #RTR_P3P4_CurrentOrder <> 0 THEN
                   #RTR_P3P4_CurrentOrder += #n;
               END_IF;


               // Transfer Pallet Roller TO Roller - PP4 TO OUTBOUND

               IF #RTR_P4TO_CurrentOrder <> 0 THEN
                   #RTR_P4TO_CurrentOrder += #n;
               END_IF;


               // Transfer Pallet Chain to Chain
               IF #Chain_To_Chain_CurrentOrder <> 0 THEN
                   #Chain_To_Chain_CurrentOrder += #n;
               END_IF;

               // Transfer TO pick station (From Pop Conveyor 4)
               IF #Pop4_To_PickSt_CurrentOrder <> 0 THEN
                   #Pop4_To_PickSt_CurrentOrder += #n;
               END_IF;

               // Transfer from Pick station (To Pop Conveyor 1)
               IF #PickSt_To_Pop1_CurrentOrder <> 0 THEN
                   #PickSt_To_Pop1_CurrentOrder += #n;
               END_IF;


               //Weigh Station
               IF #WeighingStation_CurrentOrder <> 0 THEN
                   #WeighingStation_CurrentOrder += #n;
               END_IF;

               //Profile Station
               IF #ProfileStation_CurrentOrder <> 0 THEN
                   #ProfileStation_CurrentOrder += #n;
               END_IF;


           END_IF;
            #System.OrderSent := FALSE;
       END_IF;
   END_REGION

   REGION Auto/Man Mode
       //Enable Devices in Auto/Man Mode
       IF #System.Auto_Man THEN
         //  #Cnv_Entry.Mode := #Cnv_PopUp_1.Mode:= #WeighingStation.Mode := #ProfileStation.Mode :=
          // #Cnv_PopUp_2.Mode := #Cnv_PopUp_3.Mode := #Cnv_PopUp_4.Mode := #Cnv_Exit.Mode := 3;// Auto Mode

           #Cnv_Entry.Instruction.Enable := #Cnv_PopUp_1.Instruction.Enable := #WeighingStation.Enable :=
           #ProfileStation.Enable := #Cnv_PopUp_2.Instruction.Enable := #Cnv_PopUp_3.Enabled := #Cnv_PopUp_4.Instruction.Enable :=
           #Cnv_Exit.Instruction.Enable := TRUE; // := Not System.Error

       ELSE //Disable Devices in Auto/Man Mode
          // #Cnv_Entry.Mode := #Cnv_PopUp_1.Mode := #WeighingStation.Mode := #ProfileStation.Mode :=
         //  #Cnv_PopUp_2.Mode := #Cnv_PopUp_3.Mode := #Cnv_PopUp_4.Mode := #Cnv_Exit.Mode:= 0;
           #Cnv_Entry.Instruction.Enable := #Cnv_PopUp_1.Instruction.Enable := #WeighingStation.Enable :=
           #ProfileStation.Enable := #Cnv_PopUp_2.Instruction.Enable := #Cnv_PopUp_3.Enabled := #Cnv_PopUp_4.Instruction.Enable :=
           #Cnv_Exit.Instruction.Enable := FALSE;
       END_IF;
   END_REGION

   REGION Roller to Roller - Carousel Conveyors - Original
       //Roller conveyors
       IF #System.OrderTable[1].StepNo <> 0
           AND #System.OrderTable[1].Device = #ROLLER_TO_ROLLER_DEVICE
           AND #System.OrderTable[1].Status = #QUEUED_STATUS
          // AND NOT (#Cnv_Entry.Running OR #Cnv_Exit.Running OR #Cnv_PopUp_1.Running OR #Cnv_PopUp_2.Running  OR #Cnv_PopUp_3.Running OR #Cnv_PopUp_4.Running)
           AND NOT #System.Error
           AND NOT #Canceling
         //  AND #System.OrderTable[#PickSt_To_Pop1_CurrentOrder].Status <> #RUNNING_STATUS
           //AND #System.OrderTable[#Roller_To_Roller_CurrentOrder].Status <> #RUNNING_STATUS
          // AND #System.OrderTable[#Chain_To_Chain_CurrentOrder].Status <> #RUNNING_STATUS
          // 
          // AND "OPC_UA_Control_FB_DB".State_Carrousel = 10 // OPC UA ready to receive next transaction
       THEN
           #Roller_To_Roller_CurrentOrder := 1;
       END_IF;
       IF #System.OrderTable[#Roller_To_Roller_CurrentOrder].StepNo <> 0
           AND #System.OrderTable[#Roller_To_Roller_CurrentOrder].Device = #ROLLER_TO_ROLLER_DEVICE
           AND #System.OrderTable[#Roller_To_Roller_CurrentOrder].Status = #QUEUED_STATUS
           //AND NOT (#Cnv_Entry.Running OR #Cnv_Exit.Running OR #Cnv_PopUp_1.Running OR #Cnv_PopUp_2.Running  OR #Cnv_PopUp_3.Running OR #Cnv_PopUp_4.Running)
           AND NOT #System.Error
           AND NOT #Canceling
          // AND #System.OrderTable[#PickSt_To_Pop1_CurrentOrder].Status <> #RUNNING_STATUS
          //AND #System.OrderTable[#Roller_To_Roller_CurrentOrder].Status <> #RUNNING_STATUS
          // AND #System.OrderTable[#Chain_To_Chain_CurrentOrder].Status <> #RUNNING_STATUS
       THEN
           //OPC Commands to Move Pallets - Carousel Conveyors
           // WCS => Order Table => OPC Ua Control Table
           // 
           IF #System.OrderTable[1].OPC_Control.Task_Type = 14 THEN // Profile Station - P1 TO P2
               "Control_DB"."Profiling Station".Start := TRUE;
           ELSE
               "Control_DB"."Profiling Station".Start :=FALSE;
           END_IF;

           IF #System.OrderTable[1].OPC_Control.Task_Type = 16 THEN // Barcode Scanner - INB TO P1
               "Control_DB"."InBarcode_Station".Start := TRUE;
           ELSE
               "Control_DB"."InBarcode_Station".Start := FALSE;
           END_IF;

           //"Control_DB".InBarcode_Station.Start := TRUE;
           "Control_DB"."Carrousel_Order Table".Task_Data_Available := TRUE;//#System.OrderTable[#Roller_To_Roller_CurrentOrder].OPC_Control.Task_Data_Available; // Send the Task Data Available from WCS 
           "Control_DB"."Carrousel_Order Table".Task_Type := #System.OrderTable[#Roller_To_Roller_CurrentOrder].OPC_Control.Task_Type; //  Send the Task Type - Roller to Roller Conveyor = Task Type = 6
           "Control_DB"."Carrousel_Order Table".Task_ID := #System.OrderTable[#Roller_To_Roller_CurrentOrder].OPC_Control.Task_ID; // Send the Task ID number;
           "Control_DB"."Carrousel_Order Table".Task_Metadata := #System.OrderTable[#Roller_To_Roller_CurrentOrder].OPC_Control.Task_Metadata; // Send the Task Metadata Unique identifier
           "Control_DB"."Carrousel_Order Table".Source_Location:=#System.OrderTable[#Roller_To_Roller_CurrentOrder].OPC_Control.Source_Location; // Send the Source Location from the Conveyor
           "Control_DB"."Carrousel_Order Table".Destination_Location := #System.OrderTable[#Roller_To_Roller_CurrentOrder].OPC_Control.Destination_Location; // Send the Destination Location to the Conveyor;
           #Roller_To_Roller_WatchdogStart := true;


       END_IF;

       //RUNNING
       IF (#Cnv_Entry.Running OR #Cnv_Exit.Running OR #Cnv_PopUp_1.Running OR #Cnv_PopUp_2.Running
           OR #Cnv_PopUp_3.Running OR #Cnv_PopUp_4.Running)AND #System.Auto_Man THEN
           // "Control_DB"."Profiling Station".Start := FALSE;
           // "Control_DB".InBarcode_Station.Start := FALSE;
           // "Control_DB"."Carrousel_Order Table".Task_Data_Available := FALSE; // Send the Task Data Available from WCS 
           // "Control_DB"."Carrousel_Order Table".Task_Type := 0; //  Send the Task Type - Roller to Roller Conveyor = Task Type = 6
           // "Control_DB"."Carrousel_Order Table".Task_ID := 0; // Send the Task ID number;
           // "Control_DB"."Carrousel_Order Table".Task_Metadata := ''; // Send the Task Metadata Unique identifier
           // "Control_DB"."Carrousel_Order Table".Source_Location := 0; // Send the Source Location from the Conveyor
           // "Control_DB"."Carrousel_Order Table".Destination_Location := 0; // Send the Destination Location to the Conveyor;

           //#Cnv_Entry.Instruction.Execute := FALSE;
           #System.OrderTable[#Roller_To_Roller_CurrentOrder].Status := #RUNNING_STATUS;
       END_IF;

       //Cancel order
       IF #Canceling AND NOT (#Cnv_Entry.Running OR #Cnv_Exit.Running OR #Cnv_PopUp_1.Running OR
           #Cnv_PopUp_2.Running OR #Cnv_PopUp_3.Running OR #Cnv_PopUp_4.Running) AND #Roller_To_Roller_CurrentOrder <> 0
       THEN
           #System.OrderTable[#Roller_To_Roller_CurrentOrder].Status := #CANCELED_STATUS;
           #System.OrderTable[#Roller_To_Roller_CurrentOrder].CompleteTime := #CurrentTime;
           #Roller_To_Roller_CurrentOrder := 0;

           "Control_DB"."Profiling Station".Start := FALSE;
           "Control_DB".InBarcode_Station.Start := FALSE;
           "Control_DB"."Carrousel_Order Table".Task_Data_Available := FALSE; // Send the Task Data Available from WCS 
           "Control_DB"."Carrousel_Order Table".Task_Type := 0; //  Send the Task Type - Roller to Roller Conveyor = Task Type = 6
           "Control_DB"."Carrousel_Order Table".Task_ID := 0; // Send the Task ID number;
           "Control_DB"."Carrousel_Order Table".Task_Metadata := ''; // Send the Task Metadata Unique identifier
           "Control_DB"."Carrousel_Order Table".Source_Location := 0; // Send the Source Location from the Conveyor
           "Control_DB"."Carrousel_Order Table".Destination_Location := 0; // Send the Destination Location to the Conveyor;
           //#Cnv_Entry.Instruction.Execute := FALSE;
       END_IF;

       //Error
       IF (#Cnv_Entry.Error OR #Cnv_Exit.Error OR #Cnv_PopUp_1.Error OR #Cnv_PopUp_2.Error OR #Cnv_PopUp_3.Error OR #Cnv_PopUp_4.Error) THEN
           //#Cnv_Entry.Instruction.Execute := FALSE;
           "Control_DB"."Profiling Station".Start := FALSE;
           "Control_DB".InBarcode_Station.Start := FALSE;
           "Control_DB"."Carrousel_Order Table".Task_Data_Available := FALSE; // Send the Task Data Available from WCS 
           "Control_DB"."Carrousel_Order Table".Task_Type := 0; //  Send the Task Type - Roller to Roller Conveyor = Task Type = 6
           "Control_DB"."Carrousel_Order Table".Task_ID := 0; // Send the Task ID number;
           "Control_DB"."Carrousel_Order Table".Task_Metadata := ''; // Send the Task Metadata Unique identifier
           "Control_DB"."Carrousel_Order Table".Source_Location := 0; // Send the Source Location from the Conveyor
           "Control_DB"."Carrousel_Order Table".Destination_Location := 0; // Send the Destination Location to the Conveyor;
           #System.OrderTable[#Roller_To_Roller_CurrentOrder].ErrorID := (#Cnv_Entry.Cnv_Errors.Error_Word_4
           OR #Cnv_Exit.Cnv_Errors.Error_Word_4
           OR #Cnv_PopUp_1.Cnv_Errors.Error_Word_1
           OR #Cnv_PopUp_2.Cnv_Errors.Error_Word_1
           OR #Cnv_PopUp_3.Cnv_Errors.Error_Word_1
           OR #Cnv_PopUp_4.Cnv_Errors.Error_Word_1);

       END_IF;

       //MOVEMENT FINALIZED
       #Roller_To_RollerDoneRTrig(CLK :="Control_DB"."Carrousel_Order Table".Movement_Request_Complete);
       IF #Roller_To_RollerDoneRTrig.Q THEN

           "Control_DB"."Profiling Station".Start := FALSE;
           "Control_DB".InBarcode_Station.Start := FALSE;
           "Control_DB"."Carrousel_Order Table".Task_Data_Available := FALSE; // Send the Task Data Available from WCS 
           "Control_DB"."Carrousel_Order Table".Task_Type := 0; //  Send the Task Type - Roller to Roller Conveyor = Task Type = 6
           "Control_DB"."Carrousel_Order Table".Task_ID := 0; // Send the Task ID number;
           "Control_DB"."Carrousel_Order Table".Task_Metadata := ''; // Send the Task Metadata Unique identifier
           "Control_DB"."Carrousel_Order Table".Source_Location := 0; // Send the Source Location from the Conveyor
           "Control_DB"."Carrousel_Order Table".Destination_Location := 0; // Send the Destination Location to the Conveyor;

           #Roller_To_Roller_WatchdogStart := FALSE;
           #System.OrderTable[#Roller_To_Roller_CurrentOrder].Status := #COMPLETED_STATUS;
           #System.OrderTable[#Roller_To_Roller_CurrentOrder].CompleteTime := #CurrentTime;
           #Roller_To_Roller_CurrentOrder := 0;
       END_IF;
   END_REGION

   REGION Roller TO Roller - Carousel Conveyors - Inbound to PP1 - With Barcode
   //Roller conveyors
   IF #System.OrderTable[1].StepNo <> 0
       AND #System.OrderTable[1].Device = #ROLLER_TO_ROLLER_DEVICE
       AND #System.OrderTable[1].Status = #QUEUED_STATUS
       // AND NOT (#Cnv_Entry.Running OR #Cnv_Exit.Running OR #Cnv_PopUp_1.Running OR #Cnv_PopUp_2.Running  OR #Cnv_PopUp_3.Running OR #Cnv_PopUp_4.Running)
       AND NOT #System.Error
       AND NOT #Canceling
       //  AND #System.OrderTable[#PickSt_To_Pop1_CurrentOrder].Status <> #RUNNING_STATUS
       //AND #System.OrderTable[#Roller_To_Roller_CurrentOrder].Status <> #RUNNING_STATUS
       // AND #System.OrderTable[#Chain_To_Chain_CurrentOrder].Status <> #RUNNING_STATUS
       // 
       // AND "OPC_UA_Control_FB_DB".State_Carrousel = 10 // OPC UA ready to receive next transaction
   THEN
       #Roller_To_Roller_CurrentOrder := 1;
   END_IF;
   IF #System.OrderTable[#Roller_To_Roller_CurrentOrder].StepNo <> 0
       AND #System.OrderTable[#Roller_To_Roller_CurrentOrder].Device = #ROLLER_TO_ROLLER_DEVICE
       AND #System.OrderTable[#Roller_To_Roller_CurrentOrder].Status = #QUEUED_STATUS
       //AND NOT (#Cnv_Entry.Running OR #Cnv_Exit.Running OR #Cnv_PopUp_1.Running OR #Cnv_PopUp_2.Running  OR #Cnv_PopUp_3.Running OR #Cnv_PopUp_4.Running)
       AND NOT #System.Error
       AND NOT #Canceling
       // AND #System.OrderTable[#PickSt_To_Pop1_CurrentOrder].Status <> #RUNNING_STATUS
       //AND #System.OrderTable[#Roller_To_Roller_CurrentOrder].Status <> #RUNNING_STATUS
       // AND #System.OrderTable[#Chain_To_Chain_CurrentOrder].Status <> #RUNNING_STATUS
   THEN
       //OPC Commands to Move Pallets - Carousel Conveyors
       // WCS => Order Table => OPC Ua Control Table
       // 
       IF #System.OrderTable[1].OPC_Control.Task_Type = 14 THEN // Profile Station - P1 TO P2
           "Control_DB"."Profiling Station".Start := TRUE;
       ELSE
           "Control_DB"."Profiling Station".Start := FALSE;
       END_IF;

       IF #System.OrderTable[1].OPC_Control.Task_Type = 16 THEN // Barcode Scanner - INB TO P1
           "Control_DB"."InBarcode_Station".Start := TRUE;
       ELSE
           "Control_DB"."InBarcode_Station".Start := FALSE;
       END_IF;

       //"Control_DB".InBarcode_Station.Start := TRUE;
       "Control_DB"."Carrousel_Order Table".Task_Data_Available := TRUE;//#System.OrderTable[#Roller_To_Roller_CurrentOrder].OPC_Control.Task_Data_Available; // Send the Task Data Available from WCS 
       "Control_DB"."Carrousel_Order Table".Task_Type := #System.OrderTable[#Roller_To_Roller_CurrentOrder].OPC_Control.Task_Type; //  Send the Task Type - Roller to Roller Conveyor = Task Type = 6
       "Control_DB"."Carrousel_Order Table".Task_ID := #System.OrderTable[#Roller_To_Roller_CurrentOrder].OPC_Control.Task_ID; // Send the Task ID number;
       "Control_DB"."Carrousel_Order Table".Task_Metadata := #System.OrderTable[#Roller_To_Roller_CurrentOrder].OPC_Control.Task_Metadata; // Send the Task Metadata Unique identifier
       "Control_DB"."Carrousel_Order Table".Source_Location := #System.OrderTable[#Roller_To_Roller_CurrentOrder].OPC_Control.Source_Location; // Send the Source Location from the Conveyor
       "Control_DB"."Carrousel_Order Table".Destination_Location := #System.OrderTable[#Roller_To_Roller_CurrentOrder].OPC_Control.Destination_Location; // Send the Destination Location to the Conveyor;
       #Roller_To_Roller_WatchdogStart := true;


   END_IF;

   //RUNNING
   IF (#Cnv_Entry.Running OR #Cnv_Exit.Running OR #Cnv_PopUp_1.Running OR #Cnv_PopUp_2.Running
       OR #Cnv_PopUp_3.Running OR #Cnv_PopUp_4.Running) AND #System.Auto_Man THEN
       // "Control_DB"."Profiling Station".Start := FALSE;
       // "Control_DB".InBarcode_Station.Start := FALSE;
       // "Control_DB"."Carrousel_Order Table".Task_Data_Available := FALSE; // Send the Task Data Available from WCS 
       // "Control_DB"."Carrousel_Order Table".Task_Type := 0; //  Send the Task Type - Roller to Roller Conveyor = Task Type = 6
       // "Control_DB"."Carrousel_Order Table".Task_ID := 0; // Send the Task ID number;
       // "Control_DB"."Carrousel_Order Table".Task_Metadata := ''; // Send the Task Metadata Unique identifier
       // "Control_DB"."Carrousel_Order Table".Source_Location := 0; // Send the Source Location from the Conveyor
       // "Control_DB"."Carrousel_Order Table".Destination_Location := 0; // Send the Destination Location to the Conveyor;

       //#Cnv_Entry.Instruction.Execute := FALSE;
       #System.OrderTable[#Roller_To_Roller_CurrentOrder].Status := #RUNNING_STATUS;
   END_IF;

   //Cancel order
   IF #Canceling AND NOT (#Cnv_Entry.Running OR #Cnv_Exit.Running OR #Cnv_PopUp_1.Running OR
       #Cnv_PopUp_2.Running OR #Cnv_PopUp_3.Running OR #Cnv_PopUp_4.Running) AND #Roller_To_Roller_CurrentOrder <> 0
   THEN
       #System.OrderTable[#Roller_To_Roller_CurrentOrder].Status := #CANCELED_STATUS;
       #System.OrderTable[#Roller_To_Roller_CurrentOrder].CompleteTime := #CurrentTime;
       #Roller_To_Roller_CurrentOrder := 0;

       "Control_DB"."Profiling Station".Start := FALSE;
       "Control_DB".InBarcode_Station.Start := FALSE;
       "Control_DB"."Carrousel_Order Table".Task_Data_Available := FALSE; // Send the Task Data Available from WCS 
       "Control_DB"."Carrousel_Order Table".Task_Type := 0; //  Send the Task Type - Roller to Roller Conveyor = Task Type = 6
       "Control_DB"."Carrousel_Order Table".Task_ID := 0; // Send the Task ID number;
       "Control_DB"."Carrousel_Order Table".Task_Metadata := ''; // Send the Task Metadata Unique identifier
       "Control_DB"."Carrousel_Order Table".Source_Location := 0; // Send the Source Location from the Conveyor
       "Control_DB"."Carrousel_Order Table".Destination_Location := 0; // Send the Destination Location to the Conveyor;
       //#Cnv_Entry.Instruction.Execute := FALSE;
   END_IF;

   //Error
   IF (#Cnv_Entry.Error OR #Cnv_Exit.Error OR #Cnv_PopUp_1.Error OR #Cnv_PopUp_2.Error OR #Cnv_PopUp_3.Error OR #Cnv_PopUp_4.Error) THEN
       //#Cnv_Entry.Instruction.Execute := FALSE;
       "Control_DB"."Profiling Station".Start := FALSE;
       "Control_DB".InBarcode_Station.Start := FALSE;
       "Control_DB"."Carrousel_Order Table".Task_Data_Available := FALSE; // Send the Task Data Available from WCS 
       "Control_DB"."Carrousel_Order Table".Task_Type := 0; //  Send the Task Type - Roller to Roller Conveyor = Task Type = 6
       "Control_DB"."Carrousel_Order Table".Task_ID := 0; // Send the Task ID number;
       "Control_DB"."Carrousel_Order Table".Task_Metadata := ''; // Send the Task Metadata Unique identifier
       "Control_DB"."Carrousel_Order Table".Source_Location := 0; // Send the Source Location from the Conveyor
       "Control_DB"."Carrousel_Order Table".Destination_Location := 0; // Send the Destination Location to the Conveyor;
       #System.OrderTable[#Roller_To_Roller_CurrentOrder].ErrorID := (#Cnv_Entry.Cnv_Errors.Error_Word_4
       OR #Cnv_Exit.Cnv_Errors.Error_Word_4
       OR #Cnv_PopUp_1.Cnv_Errors.Error_Word_1
       OR #Cnv_PopUp_2.Cnv_Errors.Error_Word_1
       OR #Cnv_PopUp_3.Cnv_Errors.Error_Word_1
       OR #Cnv_PopUp_4.Cnv_Errors.Error_Word_1);

   END_IF;

   //MOVEMENT FINALIZED
   #Roller_To_RollerDoneRTrig(CLK := "Control_DB"."Carrousel_Order Table".Movement_Request_Complete);
   IF #Roller_To_RollerDoneRTrig.Q THEN

       "Control_DB"."Profiling Station".Start := FALSE;
       "Control_DB".InBarcode_Station.Start := FALSE;
       "Control_DB"."Carrousel_Order Table".Task_Data_Available := FALSE; // Send the Task Data Available from WCS 
       "Control_DB"."Carrousel_Order Table".Task_Type := 0; //  Send the Task Type - Roller to Roller Conveyor = Task Type = 6
       "Control_DB"."Carrousel_Order Table".Task_ID := 0; // Send the Task ID number;
       "Control_DB"."Carrousel_Order Table".Task_Metadata := ''; // Send the Task Metadata Unique identifier
       "Control_DB"."Carrousel_Order Table".Source_Location := 0; // Send the Source Location from the Conveyor
       "Control_DB"."Carrousel_Order Table".Destination_Location := 0; // Send the Destination Location to the Conveyor;

       #Roller_To_Roller_WatchdogStart := FALSE;
       #System.OrderTable[#Roller_To_Roller_CurrentOrder].Status := #COMPLETED_STATUS;
       #System.OrderTable[#Roller_To_Roller_CurrentOrder].CompleteTime := #CurrentTime;
       #Roller_To_Roller_CurrentOrder := 0;
   END_IF;
   END_REGION

   REGION Roller TO Roller - Carousel Conveyors - PP1 to PP2 - With Profile Station
       //Roller conveyors
       IF #System.OrderTable[1].StepNo <> 0
           AND #System.OrderTable[1].Device = #ROLLER_TO_ROLLER_DEVICE
           AND #System.OrderTable[1].Status = #QUEUED_STATUS
           // AND NOT (#Cnv_Entry.Running OR #Cnv_Exit.Running OR #Cnv_PopUp_1.Running OR #Cnv_PopUp_2.Running  OR #Cnv_PopUp_3.Running OR #Cnv_PopUp_4.Running)
           AND NOT #System.Error
           AND NOT #Canceling
           //  AND #System.OrderTable[#PickSt_To_Pop1_CurrentOrder].Status <> #RUNNING_STATUS
           //AND #System.OrderTable[#Roller_To_Roller_CurrentOrder].Status <> #RUNNING_STATUS
           // AND #System.OrderTable[#Chain_To_Chain_CurrentOrder].Status <> #RUNNING_STATUS
           // 
           // AND "OPC_UA_Control_FB_DB".State_Carrousel = 10 // OPC UA ready to receive next transaction
       THEN
           #Roller_To_Roller_CurrentOrder := 1;
       END_IF;
       IF #System.OrderTable[#Roller_To_Roller_CurrentOrder].StepNo <> 0
           AND #System.OrderTable[#Roller_To_Roller_CurrentOrder].Device = #ROLLER_TO_ROLLER_DEVICE
           AND #System.OrderTable[#Roller_To_Roller_CurrentOrder].Status = #QUEUED_STATUS
           //AND NOT (#Cnv_Entry.Running OR #Cnv_Exit.Running OR #Cnv_PopUp_1.Running OR #Cnv_PopUp_2.Running  OR #Cnv_PopUp_3.Running OR #Cnv_PopUp_4.Running)
           AND NOT #System.Error
           AND NOT #Canceling
           // AND #System.OrderTable[#PickSt_To_Pop1_CurrentOrder].Status <> #RUNNING_STATUS
           //AND #System.OrderTable[#Roller_To_Roller_CurrentOrder].Status <> #RUNNING_STATUS
           // AND #System.OrderTable[#Chain_To_Chain_CurrentOrder].Status <> #RUNNING_STATUS
       THEN
           //OPC Commands to Move Pallets - Carousel Conveyors
           // WCS => Order Table => OPC Ua Control Table
           // 
           IF #System.OrderTable[1].OPC_Control.Task_Type = 14 THEN // Profile Station - P1 TO P2
               "Control_DB"."Profiling Station".Start := TRUE;
           ELSE
               "Control_DB"."Profiling Station".Start := FALSE;
           END_IF;

           IF #System.OrderTable[1].OPC_Control.Task_Type = 16 THEN // Barcode Scanner - INB TO P1
               "Control_DB"."InBarcode_Station".Start := TRUE;
           ELSE
               "Control_DB"."InBarcode_Station".Start := FALSE;
           END_IF;

           //"Control_DB".InBarcode_Station.Start := TRUE;
           "Control_DB"."Carrousel_Order Table".Task_Data_Available := TRUE;//#System.OrderTable[#Roller_To_Roller_CurrentOrder].OPC_Control.Task_Data_Available; // Send the Task Data Available from WCS 
           "Control_DB"."Carrousel_Order Table".Task_Type := #System.OrderTable[#Roller_To_Roller_CurrentOrder].OPC_Control.Task_Type; //  Send the Task Type - Roller to Roller Conveyor = Task Type = 6
           "Control_DB"."Carrousel_Order Table".Task_ID := #System.OrderTable[#Roller_To_Roller_CurrentOrder].OPC_Control.Task_ID; // Send the Task ID number;
           "Control_DB"."Carrousel_Order Table".Task_Metadata := #System.OrderTable[#Roller_To_Roller_CurrentOrder].OPC_Control.Task_Metadata; // Send the Task Metadata Unique identifier
           "Control_DB"."Carrousel_Order Table".Source_Location := #System.OrderTable[#Roller_To_Roller_CurrentOrder].OPC_Control.Source_Location; // Send the Source Location from the Conveyor
           "Control_DB"."Carrousel_Order Table".Destination_Location := #System.OrderTable[#Roller_To_Roller_CurrentOrder].OPC_Control.Destination_Location; // Send the Destination Location to the Conveyor;
           #Roller_To_Roller_WatchdogStart := true;


       END_IF;

       //RUNNING
       IF (#Cnv_Entry.Running OR #Cnv_Exit.Running OR #Cnv_PopUp_1.Running OR #Cnv_PopUp_2.Running
           OR #Cnv_PopUp_3.Running OR #Cnv_PopUp_4.Running) AND #System.Auto_Man THEN
           // "Control_DB"."Profiling Station".Start := FALSE;
           // "Control_DB".InBarcode_Station.Start := FALSE;
           // "Control_DB"."Carrousel_Order Table".Task_Data_Available := FALSE; // Send the Task Data Available from WCS 
           // "Control_DB"."Carrousel_Order Table".Task_Type := 0; //  Send the Task Type - Roller to Roller Conveyor = Task Type = 6
           // "Control_DB"."Carrousel_Order Table".Task_ID := 0; // Send the Task ID number;
           // "Control_DB"."Carrousel_Order Table".Task_Metadata := ''; // Send the Task Metadata Unique identifier
           // "Control_DB"."Carrousel_Order Table".Source_Location := 0; // Send the Source Location from the Conveyor
           // "Control_DB"."Carrousel_Order Table".Destination_Location := 0; // Send the Destination Location to the Conveyor;

           //#Cnv_Entry.Instruction.Execute := FALSE;
           #System.OrderTable[#Roller_To_Roller_CurrentOrder].Status := #RUNNING_STATUS;
       END_IF;

       //Cancel order
       IF #Canceling AND NOT (#Cnv_Entry.Running OR #Cnv_Exit.Running OR #Cnv_PopUp_1.Running OR
           #Cnv_PopUp_2.Running OR #Cnv_PopUp_3.Running OR #Cnv_PopUp_4.Running) AND #Roller_To_Roller_CurrentOrder <> 0
       THEN
           #System.OrderTable[#Roller_To_Roller_CurrentOrder].Status := #CANCELED_STATUS;
           #System.OrderTable[#Roller_To_Roller_CurrentOrder].CompleteTime := #CurrentTime;
           #Roller_To_Roller_CurrentOrder := 0;

           "Control_DB"."Profiling Station".Start := FALSE;
           "Control_DB".InBarcode_Station.Start := FALSE;
           "Control_DB"."Carrousel_Order Table".Task_Data_Available := FALSE; // Send the Task Data Available from WCS 
           "Control_DB"."Carrousel_Order Table".Task_Type := 0; //  Send the Task Type - Roller to Roller Conveyor = Task Type = 6
           "Control_DB"."Carrousel_Order Table".Task_ID := 0; // Send the Task ID number;
           "Control_DB"."Carrousel_Order Table".Task_Metadata := ''; // Send the Task Metadata Unique identifier
           "Control_DB"."Carrousel_Order Table".Source_Location := 0; // Send the Source Location from the Conveyor
           "Control_DB"."Carrousel_Order Table".Destination_Location := 0; // Send the Destination Location to the Conveyor;
           //#Cnv_Entry.Instruction.Execute := FALSE;
       END_IF;

       //Error
       IF (#Cnv_Entry.Error OR #Cnv_Exit.Error OR #Cnv_PopUp_1.Error OR #Cnv_PopUp_2.Error OR #Cnv_PopUp_3.Error OR #Cnv_PopUp_4.Error) THEN
           //#Cnv_Entry.Instruction.Execute := FALSE;
           "Control_DB"."Profiling Station".Start := FALSE;
           "Control_DB".InBarcode_Station.Start := FALSE;
           "Control_DB"."Carrousel_Order Table".Task_Data_Available := FALSE; // Send the Task Data Available from WCS 
           "Control_DB"."Carrousel_Order Table".Task_Type := 0; //  Send the Task Type - Roller to Roller Conveyor = Task Type = 6
           "Control_DB"."Carrousel_Order Table".Task_ID := 0; // Send the Task ID number;
           "Control_DB"."Carrousel_Order Table".Task_Metadata := ''; // Send the Task Metadata Unique identifier
           "Control_DB"."Carrousel_Order Table".Source_Location := 0; // Send the Source Location from the Conveyor
           "Control_DB"."Carrousel_Order Table".Destination_Location := 0; // Send the Destination Location to the Conveyor;
           #System.OrderTable[#Roller_To_Roller_CurrentOrder].ErrorID := (#Cnv_Entry.Cnv_Errors.Error_Word_4
           OR #Cnv_Exit.Cnv_Errors.Error_Word_4
           OR #Cnv_PopUp_1.Cnv_Errors.Error_Word_1
           OR #Cnv_PopUp_2.Cnv_Errors.Error_Word_1
           OR #Cnv_PopUp_3.Cnv_Errors.Error_Word_1
           OR #Cnv_PopUp_4.Cnv_Errors.Error_Word_1);

       END_IF;

       //MOVEMENT FINALIZED
       #Roller_To_RollerDoneRTrig(CLK := "Control_DB"."Carrousel_Order Table".Movement_Request_Complete);
       IF #Roller_To_RollerDoneRTrig.Q THEN

           "Control_DB"."Profiling Station".Start := FALSE;
           "Control_DB".InBarcode_Station.Start := FALSE;
           "Control_DB"."Carrousel_Order Table".Task_Data_Available := FALSE; // Send the Task Data Available from WCS 
           "Control_DB"."Carrousel_Order Table".Task_Type := 0; //  Send the Task Type - Roller to Roller Conveyor = Task Type = 6
           "Control_DB"."Carrousel_Order Table".Task_ID := 0; // Send the Task ID number;
           "Control_DB"."Carrousel_Order Table".Task_Metadata := ''; // Send the Task Metadata Unique identifier
           "Control_DB"."Carrousel_Order Table".Source_Location := 0; // Send the Source Location from the Conveyor
           "Control_DB"."Carrousel_Order Table".Destination_Location := 0; // Send the Destination Location to the Conveyor;

           #Roller_To_Roller_WatchdogStart := FALSE;
           #System.OrderTable[#Roller_To_Roller_CurrentOrder].Status := #COMPLETED_STATUS;
           #System.OrderTable[#Roller_To_Roller_CurrentOrder].CompleteTime := #CurrentTime;
           #Roller_To_Roller_CurrentOrder := 0;
       END_IF;
   END_REGION

   REGION Roller TO Roller - Carousel Conveyors - PP3 to PP4
       //Roller conveyors
       IF #System.OrderTable[1].StepNo <> 0
           AND #System.OrderTable[1].Device = #ROLLER_TO_ROLLER_DEVICE
           AND #System.OrderTable[1].Status = #QUEUED_STATUS
           // AND NOT (#Cnv_Entry.Running OR #Cnv_Exit.Running OR #Cnv_PopUp_1.Running OR #Cnv_PopUp_2.Running  OR #Cnv_PopUp_3.Running OR #Cnv_PopUp_4.Running)
           AND NOT #System.Error
           AND NOT #Canceling
           //  AND #System.OrderTable[#PickSt_To_Pop1_CurrentOrder].Status <> #RUNNING_STATUS
           //AND #System.OrderTable[#Roller_To_Roller_CurrentOrder].Status <> #RUNNING_STATUS
           // AND #System.OrderTable[#Chain_To_Chain_CurrentOrder].Status <> #RUNNING_STATUS
           // 
           // AND "OPC_UA_Control_FB_DB".State_Carrousel = 10 // OPC UA ready to receive next transaction
       THEN
           #Roller_To_Roller_CurrentOrder := 1;
       END_IF;
       IF #System.OrderTable[#Roller_To_Roller_CurrentOrder].StepNo <> 0
           AND #System.OrderTable[#Roller_To_Roller_CurrentOrder].Device = #ROLLER_TO_ROLLER_DEVICE
           AND #System.OrderTable[#Roller_To_Roller_CurrentOrder].Status = #QUEUED_STATUS
           //AND NOT (#Cnv_Entry.Running OR #Cnv_Exit.Running OR #Cnv_PopUp_1.Running OR #Cnv_PopUp_2.Running  OR #Cnv_PopUp_3.Running OR #Cnv_PopUp_4.Running)
           AND NOT #System.Error
           AND NOT #Canceling
           // AND #System.OrderTable[#PickSt_To_Pop1_CurrentOrder].Status <> #RUNNING_STATUS
           //AND #System.OrderTable[#Roller_To_Roller_CurrentOrder].Status <> #RUNNING_STATUS
           // AND #System.OrderTable[#Chain_To_Chain_CurrentOrder].Status <> #RUNNING_STATUS
       THEN
           //OPC Commands to Move Pallets - Carousel Conveyors
           // WCS => Order Table => OPC Ua Control Table
           // 
           IF #System.OrderTable[1].OPC_Control.Task_Type = 14 THEN // Profile Station - P1 TO P2
               "Control_DB"."Profiling Station".Start := TRUE;
           ELSE
               "Control_DB"."Profiling Station".Start := FALSE;
           END_IF;

           IF #System.OrderTable[1].OPC_Control.Task_Type = 16 THEN // Barcode Scanner - INB TO P1
               "Control_DB"."InBarcode_Station".Start := TRUE;
           ELSE
               "Control_DB"."InBarcode_Station".Start := FALSE;
           END_IF;

           //"Control_DB".InBarcode_Station.Start := TRUE;
           "Control_DB"."Carrousel_Order Table".Task_Data_Available := TRUE;//#System.OrderTable[#Roller_To_Roller_CurrentOrder].OPC_Control.Task_Data_Available; // Send the Task Data Available from WCS 
           "Control_DB"."Carrousel_Order Table".Task_Type := #System.OrderTable[#Roller_To_Roller_CurrentOrder].OPC_Control.Task_Type; //  Send the Task Type - Roller to Roller Conveyor = Task Type = 6
           "Control_DB"."Carrousel_Order Table".Task_ID := #System.OrderTable[#Roller_To_Roller_CurrentOrder].OPC_Control.Task_ID; // Send the Task ID number;
           "Control_DB"."Carrousel_Order Table".Task_Metadata := #System.OrderTable[#Roller_To_Roller_CurrentOrder].OPC_Control.Task_Metadata; // Send the Task Metadata Unique identifier
           "Control_DB"."Carrousel_Order Table".Source_Location := #System.OrderTable[#Roller_To_Roller_CurrentOrder].OPC_Control.Source_Location; // Send the Source Location from the Conveyor
           "Control_DB"."Carrousel_Order Table".Destination_Location := #System.OrderTable[#Roller_To_Roller_CurrentOrder].OPC_Control.Destination_Location; // Send the Destination Location to the Conveyor;
           #Roller_To_Roller_WatchdogStart := true;


       END_IF;

       //RUNNING
       IF (#Cnv_Entry.Running OR #Cnv_Exit.Running OR #Cnv_PopUp_1.Running OR #Cnv_PopUp_2.Running
           OR #Cnv_PopUp_3.Running OR #Cnv_PopUp_4.Running) AND #System.Auto_Man THEN
           // "Control_DB"."Profiling Station".Start := FALSE;
           // "Control_DB".InBarcode_Station.Start := FALSE;
           // "Control_DB"."Carrousel_Order Table".Task_Data_Available := FALSE; // Send the Task Data Available from WCS 
           // "Control_DB"."Carrousel_Order Table".Task_Type := 0; //  Send the Task Type - Roller to Roller Conveyor = Task Type = 6
           // "Control_DB"."Carrousel_Order Table".Task_ID := 0; // Send the Task ID number;
           // "Control_DB"."Carrousel_Order Table".Task_Metadata := ''; // Send the Task Metadata Unique identifier
           // "Control_DB"."Carrousel_Order Table".Source_Location := 0; // Send the Source Location from the Conveyor
           // "Control_DB"."Carrousel_Order Table".Destination_Location := 0; // Send the Destination Location to the Conveyor;

           //#Cnv_Entry.Instruction.Execute := FALSE;
           #System.OrderTable[#Roller_To_Roller_CurrentOrder].Status := #RUNNING_STATUS;
       END_IF;

       //Cancel order
       IF #Canceling AND NOT (#Cnv_Entry.Running OR #Cnv_Exit.Running OR #Cnv_PopUp_1.Running OR
           #Cnv_PopUp_2.Running OR #Cnv_PopUp_3.Running OR #Cnv_PopUp_4.Running) AND #Roller_To_Roller_CurrentOrder <> 0
       THEN
           #System.OrderTable[#Roller_To_Roller_CurrentOrder].Status := #CANCELED_STATUS;
           #System.OrderTable[#Roller_To_Roller_CurrentOrder].CompleteTime := #CurrentTime;
           #Roller_To_Roller_CurrentOrder := 0;

           "Control_DB"."Profiling Station".Start := FALSE;
           "Control_DB".InBarcode_Station.Start := FALSE;
           "Control_DB"."Carrousel_Order Table".Task_Data_Available := FALSE; // Send the Task Data Available from WCS 
           "Control_DB"."Carrousel_Order Table".Task_Type := 0; //  Send the Task Type - Roller to Roller Conveyor = Task Type = 6
           "Control_DB"."Carrousel_Order Table".Task_ID := 0; // Send the Task ID number;
           "Control_DB"."Carrousel_Order Table".Task_Metadata := ''; // Send the Task Metadata Unique identifier
           "Control_DB"."Carrousel_Order Table".Source_Location := 0; // Send the Source Location from the Conveyor
           "Control_DB"."Carrousel_Order Table".Destination_Location := 0; // Send the Destination Location to the Conveyor;
           //#Cnv_Entry.Instruction.Execute := FALSE;
       END_IF;

       //Error
       IF (#Cnv_Entry.Error OR #Cnv_Exit.Error OR #Cnv_PopUp_1.Error OR #Cnv_PopUp_2.Error OR #Cnv_PopUp_3.Error OR #Cnv_PopUp_4.Error) THEN
           //#Cnv_Entry.Instruction.Execute := FALSE;
           "Control_DB"."Profiling Station".Start := FALSE;
           "Control_DB".InBarcode_Station.Start := FALSE;
           "Control_DB"."Carrousel_Order Table".Task_Data_Available := FALSE; // Send the Task Data Available from WCS 
           "Control_DB"."Carrousel_Order Table".Task_Type := 0; //  Send the Task Type - Roller to Roller Conveyor = Task Type = 6
           "Control_DB"."Carrousel_Order Table".Task_ID := 0; // Send the Task ID number;
           "Control_DB"."Carrousel_Order Table".Task_Metadata := ''; // Send the Task Metadata Unique identifier
           "Control_DB"."Carrousel_Order Table".Source_Location := 0; // Send the Source Location from the Conveyor
           "Control_DB"."Carrousel_Order Table".Destination_Location := 0; // Send the Destination Location to the Conveyor;
           #System.OrderTable[#Roller_To_Roller_CurrentOrder].ErrorID := (#Cnv_Entry.Cnv_Errors.Error_Word_4
           OR #Cnv_Exit.Cnv_Errors.Error_Word_4
           OR #Cnv_PopUp_1.Cnv_Errors.Error_Word_1
           OR #Cnv_PopUp_2.Cnv_Errors.Error_Word_1
           OR #Cnv_PopUp_3.Cnv_Errors.Error_Word_1
           OR #Cnv_PopUp_4.Cnv_Errors.Error_Word_1);

       END_IF;

       //MOVEMENT FINALIZED
       #Roller_To_RollerDoneRTrig(CLK := "Control_DB"."Carrousel_Order Table".Movement_Request_Complete);
       IF #Roller_To_RollerDoneRTrig.Q THEN

           "Control_DB"."Profiling Station".Start := FALSE;
           "Control_DB".InBarcode_Station.Start := FALSE;
           "Control_DB"."Carrousel_Order Table".Task_Data_Available := FALSE; // Send the Task Data Available from WCS 
           "Control_DB"."Carrousel_Order Table".Task_Type := 0; //  Send the Task Type - Roller to Roller Conveyor = Task Type = 6
           "Control_DB"."Carrousel_Order Table".Task_ID := 0; // Send the Task ID number;
           "Control_DB"."Carrousel_Order Table".Task_Metadata := ''; // Send the Task Metadata Unique identifier
           "Control_DB"."Carrousel_Order Table".Source_Location := 0; // Send the Source Location from the Conveyor
           "Control_DB"."Carrousel_Order Table".Destination_Location := 0; // Send the Destination Location to the Conveyor;

           #Roller_To_Roller_WatchdogStart := FALSE;
           #System.OrderTable[#Roller_To_Roller_CurrentOrder].Status := #COMPLETED_STATUS;
           #System.OrderTable[#Roller_To_Roller_CurrentOrder].CompleteTime := #CurrentTime;
           #Roller_To_Roller_CurrentOrder := 0;
       END_IF;
   END_REGION

   REGION Roller TO Roller - Carousel Conveyors - PP4 to Outbound
       //Roller conveyors
       IF #System.OrderTable[1].StepNo <> 0
           AND #System.OrderTable[1].Device = #ROLLER_TO_ROLLER_DEVICE
           AND #System.OrderTable[1].Status = #QUEUED_STATUS
           // AND NOT (#Cnv_Entry.Running OR #Cnv_Exit.Running OR #Cnv_PopUp_1.Running OR #Cnv_PopUp_2.Running  OR #Cnv_PopUp_3.Running OR #Cnv_PopUp_4.Running)
           AND NOT #System.Error
           AND NOT #Canceling
           //  AND #System.OrderTable[#PickSt_To_Pop1_CurrentOrder].Status <> #RUNNING_STATUS
           //AND #System.OrderTable[#Roller_To_Roller_CurrentOrder].Status <> #RUNNING_STATUS
           // AND #System.OrderTable[#Chain_To_Chain_CurrentOrder].Status <> #RUNNING_STATUS
           // 
           // AND "OPC_UA_Control_FB_DB".State_Carrousel = 10 // OPC UA ready to receive next transaction
       THEN
           #Roller_To_Roller_CurrentOrder := 1;
       END_IF;
       IF #System.OrderTable[#Roller_To_Roller_CurrentOrder].StepNo <> 0
           AND #System.OrderTable[#Roller_To_Roller_CurrentOrder].Device = #ROLLER_TO_ROLLER_DEVICE
           AND #System.OrderTable[#Roller_To_Roller_CurrentOrder].Status = #QUEUED_STATUS
           //AND NOT (#Cnv_Entry.Running OR #Cnv_Exit.Running OR #Cnv_PopUp_1.Running OR #Cnv_PopUp_2.Running  OR #Cnv_PopUp_3.Running OR #Cnv_PopUp_4.Running)
           AND NOT #System.Error
           AND NOT #Canceling
           // AND #System.OrderTable[#PickSt_To_Pop1_CurrentOrder].Status <> #RUNNING_STATUS
           //AND #System.OrderTable[#Roller_To_Roller_CurrentOrder].Status <> #RUNNING_STATUS
           // AND #System.OrderTable[#Chain_To_Chain_CurrentOrder].Status <> #RUNNING_STATUS
       THEN
           //OPC Commands to Move Pallets - Carousel Conveyors
           // WCS => Order Table => OPC Ua Control Table
           // 
           IF #System.OrderTable[1].OPC_Control.Task_Type = 14 THEN // Profile Station - P1 TO P2
               "Control_DB"."Profiling Station".Start := TRUE;
           ELSE
               "Control_DB"."Profiling Station".Start := FALSE;
           END_IF;

           IF #System.OrderTable[1].OPC_Control.Task_Type = 16 THEN // Barcode Scanner - INB TO P1
               "Control_DB"."InBarcode_Station".Start := TRUE;
           ELSE
               "Control_DB"."InBarcode_Station".Start := FALSE;
           END_IF;

           //"Control_DB".InBarcode_Station.Start := TRUE;
           "Control_DB"."Carrousel_Order Table".Task_Data_Available := TRUE;//#System.OrderTable[#Roller_To_Roller_CurrentOrder].OPC_Control.Task_Data_Available; // Send the Task Data Available from WCS 
           "Control_DB"."Carrousel_Order Table".Task_Type := #System.OrderTable[#Roller_To_Roller_CurrentOrder].OPC_Control.Task_Type; //  Send the Task Type - Roller to Roller Conveyor = Task Type = 6
           "Control_DB"."Carrousel_Order Table".Task_ID := #System.OrderTable[#Roller_To_Roller_CurrentOrder].OPC_Control.Task_ID; // Send the Task ID number;
           "Control_DB"."Carrousel_Order Table".Task_Metadata := #System.OrderTable[#Roller_To_Roller_CurrentOrder].OPC_Control.Task_Metadata; // Send the Task Metadata Unique identifier
           "Control_DB"."Carrousel_Order Table".Source_Location := #System.OrderTable[#Roller_To_Roller_CurrentOrder].OPC_Control.Source_Location; // Send the Source Location from the Conveyor
           "Control_DB"."Carrousel_Order Table".Destination_Location := #System.OrderTable[#Roller_To_Roller_CurrentOrder].OPC_Control.Destination_Location; // Send the Destination Location to the Conveyor;
           #Roller_To_Roller_WatchdogStart := true;


       END_IF;

       //RUNNING
       IF (#Cnv_Entry.Running OR #Cnv_Exit.Running OR #Cnv_PopUp_1.Running OR #Cnv_PopUp_2.Running
           OR #Cnv_PopUp_3.Running OR #Cnv_PopUp_4.Running) AND #System.Auto_Man THEN
           // "Control_DB"."Profiling Station".Start := FALSE;
           // "Control_DB".InBarcode_Station.Start := FALSE;
           // "Control_DB"."Carrousel_Order Table".Task_Data_Available := FALSE; // Send the Task Data Available from WCS 
           // "Control_DB"."Carrousel_Order Table".Task_Type := 0; //  Send the Task Type - Roller to Roller Conveyor = Task Type = 6
           // "Control_DB"."Carrousel_Order Table".Task_ID := 0; // Send the Task ID number;
           // "Control_DB"."Carrousel_Order Table".Task_Metadata := ''; // Send the Task Metadata Unique identifier
           // "Control_DB"."Carrousel_Order Table".Source_Location := 0; // Send the Source Location from the Conveyor
           // "Control_DB"."Carrousel_Order Table".Destination_Location := 0; // Send the Destination Location to the Conveyor;

           //#Cnv_Entry.Instruction.Execute := FALSE;
           #System.OrderTable[#Roller_To_Roller_CurrentOrder].Status := #RUNNING_STATUS;
       END_IF;

       //Cancel order
       IF #Canceling AND NOT (#Cnv_Entry.Running OR #Cnv_Exit.Running OR #Cnv_PopUp_1.Running OR
           #Cnv_PopUp_2.Running OR #Cnv_PopUp_3.Running OR #Cnv_PopUp_4.Running) AND #Roller_To_Roller_CurrentOrder <> 0
       THEN
           #System.OrderTable[#Roller_To_Roller_CurrentOrder].Status := #CANCELED_STATUS;
           #System.OrderTable[#Roller_To_Roller_CurrentOrder].CompleteTime := #CurrentTime;
           #Roller_To_Roller_CurrentOrder := 0;

           "Control_DB"."Profiling Station".Start := FALSE;
           "Control_DB".InBarcode_Station.Start := FALSE;
           "Control_DB"."Carrousel_Order Table".Task_Data_Available := FALSE; // Send the Task Data Available from WCS 
           "Control_DB"."Carrousel_Order Table".Task_Type := 0; //  Send the Task Type - Roller to Roller Conveyor = Task Type = 6
           "Control_DB"."Carrousel_Order Table".Task_ID := 0; // Send the Task ID number;
           "Control_DB"."Carrousel_Order Table".Task_Metadata := ''; // Send the Task Metadata Unique identifier
           "Control_DB"."Carrousel_Order Table".Source_Location := 0; // Send the Source Location from the Conveyor
           "Control_DB"."Carrousel_Order Table".Destination_Location := 0; // Send the Destination Location to the Conveyor;
           //#Cnv_Entry.Instruction.Execute := FALSE;
       END_IF;

       //Error
       IF (#Cnv_Entry.Error OR #Cnv_Exit.Error OR #Cnv_PopUp_1.Error OR #Cnv_PopUp_2.Error OR #Cnv_PopUp_3.Error OR #Cnv_PopUp_4.Error) THEN
           //#Cnv_Entry.Instruction.Execute := FALSE;
           "Control_DB"."Profiling Station".Start := FALSE;
           "Control_DB".InBarcode_Station.Start := FALSE;
           "Control_DB"."Carrousel_Order Table".Task_Data_Available := FALSE; // Send the Task Data Available from WCS 
           "Control_DB"."Carrousel_Order Table".Task_Type := 0; //  Send the Task Type - Roller to Roller Conveyor = Task Type = 6
           "Control_DB"."Carrousel_Order Table".Task_ID := 0; // Send the Task ID number;
           "Control_DB"."Carrousel_Order Table".Task_Metadata := ''; // Send the Task Metadata Unique identifier
           "Control_DB"."Carrousel_Order Table".Source_Location := 0; // Send the Source Location from the Conveyor
           "Control_DB"."Carrousel_Order Table".Destination_Location := 0; // Send the Destination Location to the Conveyor;
           #System.OrderTable[#Roller_To_Roller_CurrentOrder].ErrorID := (#Cnv_Entry.Cnv_Errors.Error_Word_4
           OR #Cnv_Exit.Cnv_Errors.Error_Word_4
           OR #Cnv_PopUp_1.Cnv_Errors.Error_Word_1
           OR #Cnv_PopUp_2.Cnv_Errors.Error_Word_1
           OR #Cnv_PopUp_3.Cnv_Errors.Error_Word_1
           OR #Cnv_PopUp_4.Cnv_Errors.Error_Word_1);

       END_IF;

       //MOVEMENT FINALIZED
       #Roller_To_RollerDoneRTrig(CLK := "Control_DB"."Carrousel_Order Table".Movement_Request_Complete);
       IF #Roller_To_RollerDoneRTrig.Q THEN

           "Control_DB"."Profiling Station".Start := FALSE;
           "Control_DB".InBarcode_Station.Start := FALSE;
           "Control_DB"."Carrousel_Order Table".Task_Data_Available := FALSE; // Send the Task Data Available from WCS 
           "Control_DB"."Carrousel_Order Table".Task_Type := 0; //  Send the Task Type - Roller to Roller Conveyor = Task Type = 6
           "Control_DB"."Carrousel_Order Table".Task_ID := 0; // Send the Task ID number;
           "Control_DB"."Carrousel_Order Table".Task_Metadata := ''; // Send the Task Metadata Unique identifier
           "Control_DB"."Carrousel_Order Table".Source_Location := 0; // Send the Source Location from the Conveyor
           "Control_DB"."Carrousel_Order Table".Destination_Location := 0; // Send the Destination Location to the Conveyor;

           #Roller_To_Roller_WatchdogStart := FALSE;
           #System.OrderTable[#Roller_To_Roller_CurrentOrder].Status := #COMPLETED_STATUS;
           #System.OrderTable[#Roller_To_Roller_CurrentOrder].CompleteTime := #CurrentTime;
           #Roller_To_Roller_CurrentOrder := 0;
       END_IF;
   END_REGION

   REGION Chain to Chain - Carousel Conveyors - Pop 2 to Pop 3
       IF #System.OrderTable[1].StepNo <> 0
           AND #System.OrderTable[1].Device = #CHAIN_TO_CHAIN_DEVICE
           AND #System.OrderTable[1].Status = #QUEUED_STATUS
           AND NOT (#Cnv_PopUp_2.Running OR #Cnv_PopUp_3.Running)
           AND NOT #System.Error
           AND NOT #Canceling
           AND #System.OrderTable[#Roller_To_Roller_CurrentOrder].Status <> #RUNNING_STATUS

       THEN
           #Chain_To_Chain_CurrentOrder := 1;
       END_IF;
       IF #System.OrderTable[#Chain_To_Chain_CurrentOrder].StepNo <> 0
           AND #System.OrderTable[#Chain_To_Chain_CurrentOrder].Device = #CHAIN_TO_CHAIN_DEVICE
           AND #System.OrderTable[#Chain_To_Chain_CurrentOrder].Status = #QUEUED_STATUS
           AND NOT (#Cnv_PopUp_2.Running OR #Cnv_PopUp_3.Running)
           AND NOT #System.Error
           AND NOT #Canceling
           AND #System.OrderTable[#Roller_To_Roller_CurrentOrder].Status <> #RUNNING_STATUS
       THEN
           //OPC Commands to Move Pallets - Carousel Conveyors
           // WCS => Order Table => OPC Ua Control Table

           "Control_DB"."Carrousel_Order Table".Task_Data_Available := TRUE;//#System.OrderTable[#Chain_To_Chain_CurrentOrder].OPC_Control.Task_Data_Available; // Send the Task Data Available from WCS 
           "Control_DB"."Carrousel_Order Table".Task_Type := #System.OrderTable[#Chain_To_Chain_CurrentOrder].OPC_Control.Task_Type; //  Send the Task Type - Chain to Chain Conveyor = Task Type = 7
           "Control_DB"."Carrousel_Order Table".Task_ID := #System.OrderTable[#Chain_To_Chain_CurrentOrder].OPC_Control.Task_ID; // Send the Task ID number;
           "Control_DB"."Carrousel_Order Table".Task_Metadata := #System.OrderTable[#Chain_To_Chain_CurrentOrder].OPC_Control.Task_Metadata; // Send the Task Metadata Unique identifier
           "Control_DB"."Carrousel_Order Table".Source_Location := #System.OrderTable[#Chain_To_Chain_CurrentOrder].OPC_Control.Source_Location; // Send the Source Location from the Conveyor
           "Control_DB"."Carrousel_Order Table".Destination_Location := #System.OrderTable[#Chain_To_Chain_CurrentOrder].OPC_Control.Destination_Location; // Send the Destination Location to the Conveyor;
           #Chain_To_Chain_WatchdogStart := true;


       END_IF;

       //RUNNING
       IF (#Cnv_PopUp_2.Running OR #Cnv_PopUp_3.Running)AND #System.Auto_Man THEN
           //#Cnv_Entry.Instruction.Execute := FALSE;
           #System.OrderTable[#Chain_To_Chain_CurrentOrder].Status := #RUNNING_STATUS;
       END_IF;

       //Cancel order
       IF #Canceling AND NOT (#Cnv_PopUp_2.Running OR #Cnv_PopUp_3.Running) AND #Chain_To_Chain_CurrentOrder <> 0 THEN


           "Control_DB"."Carrousel_Order Table".Task_Data_Available := FALSE;//#System.OrderTable[#Chain_To_Chain_CurrentOrder].OPC_Control.Task_Data_Available; // Send the Task Data Available from WCS 
           "Control_DB"."Carrousel_Order Table".Task_Type := 0; //  Send the Task Type - Chain to Chain Conveyor = Task Type = 7
           "Control_DB"."Carrousel_Order Table".Task_ID := 0; // Send the Task ID number;
           "Control_DB"."Carrousel_Order Table".Task_Metadata := ''; // Send the Task Metadata Unique identifier
           "Control_DB"."Carrousel_Order Table".Source_Location := 0; // Send the Source Location from the Conveyor
           "Control_DB"."Carrousel_Order Table".Destination_Location := 0; // Send the Destination Location to the Conveyor;

